(* IEC 61131-3 sources: daoli-st-library/DL_Device (part 44) *)

(* ---- FB_DL_ValveStictionDetect.st ---- *)
(*==============================================================================
 * 组件名称 (Component)  : FB_DL_ValveStictionDetect
 * 所属子库 (Sublibrary) : DL_Device
 * 当前版本 (Version)    : 1.0.1
 * 兼容性   (Platform)   : CODESYS 3.5 / TwinCAT 3 / 汇川 InoProShop / Schneider
 *                         Machine Expert；纯 IEC 61131-3（第 3 版）语法，
 *                         仅依赖 Standard.library（R_TRIG / TON）
 * 组件分类 (Category)   : 功能块（FUNCTION_BLOCK）· 设备本体退化诊断 · 阀门黏滞
 * 功能描述 (Function)   : 用**常规运行数据**（指令 OP 与阀位 PV，无需激励试验）
 *                         在线判阀门黏滞，输出黏滞等级、黏滞带估计、方向性滞后
 *                         归一指标与停滞事件计数，并把「需要维护」语义交给
 *                         NE107 的 eMaintenanceReq。
 * 三条判据 (Criteria)   : 三条判据**并发**，缺一不升级（这是本件的核心裁定）：
 *                         (a) 方向性滞后：上升行程与下降行程在同一 OP 处 PV 之差，
 *                             即黏滞带 fDeadbandEst；
 *                         (b) 停滞拍：|ΔOP| > fStallThr 而 |ΔPV| < fMoveThr，持续
 *                             tStallTime 判一次停滞事件；
 *                         (c) 反转确认延迟：方向反转后到 PV 开始移动的时间超过
 *                             tReverseTime 判一次反转超时。
 *                         只有 (a) 超限而 (b)(c) 均无证据时，等级封顶在 eSlight
 *                         ——单个指标越限不足以判重度黏滞，这是文献反复强调的
 *                         「无单一方法 100% 可信」在本件的落地方式。
 * 等级映射 (Levels)     : eNone(0) → eOk；eSlight(10) / eModerate(20) →
 *                         eMaintenanceReq；eSevere(30) → eOutOfSpec。
 *                         黏滞是**退化**不是失效：阀门仍在调节，只是品质下降，
 *                         故最高只到 eOutOfSpec，绝不进 eFailure（故障只来自
 *                         参数非法与非有限输入）。
 * 边界声明 (Limits)     : ① **不做互相关**：需要长窗 FFT，违 O(1) 内存纪律；
 *                         ② **不做椭圆拟合**：需要二维迭代，不可逐拍复算；
 *                         ③ 输出是**趋势判据，不是黏滞量的计量级量化**——按
 *                         行业文献口径，黏滞带估计只用于纵向趋势比较与维护
 *                         排序，不可作为验收数据；④ 不替代定位器自诊断，
 *                         不做任何补偿（补偿属定位器或 APC 层职责）；
 *                         ⑤ **判据 (a) 只取准静态反转点**：同一 OP 处比较要求
 *                         前后反转点的指令差 ≤ fDeadbandMax。全行程单向斜坡
 *                         （0→100→0）的反转点 OP 差达全量程，本件不出滞后样本，
 *                         黏滞带保持 0、等级保持 eNone —— 这是**刻意的保守方向**：
 *                         在持续运动的阀上做同 OP 差分会把「纯跟随滞后」误算成
 *                         黏滞（滞后 0.3 % 会产出 0.6 % 的假黏滞带），文献明确
 *                         该法只在准静态与小幅往复下可信。需要全行程评估时应在
 *                         工艺上安排往复小步激励，或改看定位器自诊断。
 * 段序 (Cycle order)   : 段 1 默认值与单拍预清零 → 段 2 首扫初始化 →
 *                         段 3 参数闸门 → 段 4 定时器与边沿无条件刷新 →
 *                         段 5 输入域检查与快照 → 段 6 复位通道与故障锁存
 *                         （**CASE 前置，且不做状态赋值**）→ 段 7 相位机 →
 *                         段 8 采样采集 → 段 9 分析计算 → 段 10 发布与窗口重建
 *                         （含本拍复验）→ 段 11 出口钳位与保持重写 → 段 12 码位链。
 * 镜像量清单 (R38)      : `_bPosValidSnap` —— 窗口关闭那一刻的反馈有效性快照，
 *                         **唯一消费点**是段 9 的「窗口合法性闸门」；实时量
 *                         `bPosValid` 的三处消费点各自独立且不含边界量含义：
 *                         段 4 的定时器输入、段 7 的挂起迁移、段 10 的本拍复验。
 *                         窗口内的 OP/PV 一律取 `_afOpWin` / `_afPvWin` 缓存，
 *                         **绝不**在分析相读实时 `fPos` —— 这是 R38/R42 的正解。
 * 定时器清单 (R40)      : 实例名 / IN 表达式 / 断输入拍标志 / 自清位置
 *                         fbWindowWatch  / 相位为采集 AND NOT _bWindowBreak
 *                                        / _bWindowBreak / 段 4 调用后自清
 *                         fbSampleWatch  / 相位为采集 AND NOT _bSampleBreak
 *                                        / _bSampleBreak / 段 4 调用后自清，采样后置位
 *                         fbStallWatch   / 停滞条件 AND NOT _bStallBreak
 *                                        / _bStallBreak / 段 4 调用后自清
 *                         fbReverseWatch / 反转待确认 AND NOT _bReverseBreak
 *                                        / _bReverseBreak / 段 4 调用后自清
 *                         fbSinceWatch   / NOT _bSinceBreak / _bSinceBreak
 *                                        / 段 4 调用后自清，停滞事件时置位
 * 单拍标志清单 (R25)    : `_bResetPulse` 预清段 1 / 置位段 6 / 消费段 6；
 *                         `_bWindowBreak` `_bSampleBreak` `_bStallBreak`
 *                         `_bReverseBreak` `_bSinceBreak` 预清处不设（就地置位
 *                         后段 4 自清），置位点见定时器清单；
 *                         `_bStallEvent` `_bRevEvent` 预清段 1 / 置位段 8 /
 *                         消费段 8 与段 9。
 * 保持位清单 (R27)      : `_eLevel`（等级）、`_fDbHeld`（黏滞带）、`_uStallCount`
 *                         （停滞计数）、`_bSuspectHeld`（嫌疑位）四个保持量，全部
 *                         由段 11 每拍重写出口；复位沿清除（R27 的反面：复位是
 *                         保持量的唯一清除通道）。
 * 三元一致表 (R35)      : 量 / 守卫封顶 / 判据运算符
 *                         fDeadbandMax      / 钳到 ≥0.5   / 等级判据用 >=
 *                         fDeadbandModerate / 钳到 < Max  / 等级判据用 >=
 *                         轻微下限（Max 的 1/4）/ 钳到 ≥0.1 / 等级判据用 >=
 * 验收向量 (Acceptance) :
 *   V1 正常阀：OP 斜坡 0→100、PV 滞后 0.3% → eStiction=eNone、黏滞带约 0.3、
 *      停滞计数 0
 *   V2 黏滞阀：OP 每 2 s 步进 2%、PV 每 4 s 跳 3% → 三判据全成立 →
 *      eStiction=eSevere、停滞计数 ≥2、eHealth=eOutOfSpec
 *   V3（V-C 跨相复验）：分析相已缓存样本 → 判定相当拍 bPosValid 置 FALSE →
 *      **必须不发布新等级**（保持上次值 + 015D），不得用缓存样本直接出结论
 *   V4（V-D 恢复首拍）：挂起恢复后样本数从 0 重建（R41），重建窗**不发布**
 *      任何等级（比「不判 Severe」更严），只置 015C
 *   V5（V-A 域外）：fCmd 为 NaN → 031D 锁存，黏滞带保持上次值并夹进 0~100（R43）
 * 规格偏离 (Deviation)  :
 *   ① 规格未给采样周期。本件按「窗口长度 ÷ 最少样本数」推导采样周期并钳进
 *      20 ms~5 s，使一个标准窗恰好采到 nMinSamples 个样本；若窗口内样本数
 *      先达缓冲上限（128）则提前进入分析相，避免溢出。
 *   ② 规格的 eNone/eSlight 分界未给阈值。本件取「中限的 1/4」作为轻微下限
 *      （默认 2.0 × 0.25 = 0.5%），并在三元一致表中登记，避免出现无闸门的
 *      隐式阈值。
 *   ③ 规格 V4 要求「恢复首拍不得判 eSevere」。本件实现为**重建窗不发布任何
 *      等级**（只置 015C 保持上次值），比规格更严，且不引入「部分发布」的
 *      半可信语义。
 * 开源溯源 (Origin)     : 来源标签 namur-ne107 / stiction-diag / asset-health。
 *                         原创 clean-room 实现。NE107（公开推荐规范）仅提供
 *                         健康分级语义；阀黏滞的**判据思想**（方向性滞后、
 *                         停滞拍、反转确认延迟）来自控制工程公开文献的通行
 *                         定性描述，属公有领域方法学思想，不构成代码版权标的；
 *                         本件未复制任何文献代码或开源工程源码，缓冲区结构、
 *                         阈值口径、等级仲裁、状态机与全部码位 100% 本库独立
 *                         设计。T3 定位：文献仅作立项理由，不作为实现依据。
 * 修订历史 (Revision)   :
 *   2026-11-15  v1.0.0  首版入库（R13 · 泳道 A · 阀门黏滞在线诊断）
 *   2026-11-16  v1.0.1  终审修复一处、留档一处：① 距上次停滞定时器的 PT
 *                       由裸 `T#24H` 改为常量 DL_SINCE_MAX（无魔法数红线）；
 *                       ② 头注释补边界 ⑤，明确判据 (a) 在全行程单向斜坡下不出
 *                       样本的保守语义与理由（原实现无此声明，易被误读为漏判缺陷）。
 *============================================================================*)

(*-----------------------------------------------------------------------------
 * 枚举: E_DL_StictionLevel（归属本功能块，同文件发布）
 * 含义: 黏滞严重度。0 起步长 10，便于后续插入细分等级。
 *-----------------------------------------------------------------------------*)
TYPE E_DL_StictionLevel :
(
    eNone     := 0,    // 无黏滞：滞后在噪声带内 / No stiction, hysteresis within the noise band
    eSlight   := 10,   // 轻微：可察觉但影响可忽略 / Slight, noticeable but negligible
    eModerate := 20,   // 中度：调节品质下降，排入维护计划 / Moderate, control quality degraded
    eSevere   := 30    // 重度：明显黏滑运动，须尽快处理 / Severe, stick-slip motion
);
END_TYPE

(*-----------------------------------------------------------------------------
 * 枚举: E_DL_StictionPhase（归属本功能块，同文件发布）
 * 含义: 诊断相位。每个成员在段 7 有且仅有一个 CASE 标签，ELSE 只接脏值。
 *-----------------------------------------------------------------------------*)
TYPE E_DL_StictionPhase :
(
    eIdle    := 0,     // 待机：未使能或参数未通过 / Idle, disabled or parameters not accepted
    eCollect := 10,    // 采集：按采样周期入缓冲 / Collect, samples enter the ring buffer
    eAnalyze := 20,    // 分析：仅在窗口关闭当拍执行一次 / Analyze, executed once when the window closes
    eVerdict := 30,    // 判定：本拍复验后发布，再回采集 / Verdict, re-verify then publish
    eSuspend := 40,    // 挂起：反馈失效，非故障；恢复后窗口重建 / Suspended, not a fault
    eFault   := 99     // 故障：参数非法或输入非有限，锁存待复位 / Fault, latched until reset
);
END_TYPE

FUNCTION_BLOCK FB_DL_ValveStictionDetect
VAR_INPUT
    bEnable          : BOOL;                          // 使能，FALSE 时窗口冻结 [-] / Enable, freezes the window
    bReset           : BOOL;                          // 复位锁存与统计，上升沿有效 [-] / Rising edge resets latch and statistics
    fCmd             : REAL;                          // 阀门指令 OP [%]，范围 0~100 / Valve command in percent
    fPos             : REAL;                          // 阀位反馈 PV [%]，范围 0~100 / Valve position feedback in percent
    bPosValid        : BOOL := TRUE;                  // 反馈有效性，FALSE 时诊断挂起（非故障）[-] / Feedback validity, FALSE suspends
    fMoveThr         : REAL := 0.5;                   // 判阀位在动的位移阈 [%]，范围 0.1~5.0 / Movement threshold
    fStallThr        : REAL := 1.0;                   // 判指令在变的变化阈 [%]，范围 0.2~10.0 / Command change threshold
    tStallTime       : TIME := T#2S;                  // 停滞持续判据 [毫秒]，范围 100 ms~60 s / Stall duration
    tReverseTime     : TIME := T#1S;                  // 反转确认允许延迟 [毫秒]，范围 100 ms~30 s / Reverse confirmation delay
    tWindow          : TIME := T#60S;                 // 分析窗长 [毫秒]，范围 10 s~30 min / Analysis window
    nMinSamples      : INT := 30;                     // 窗口最少有效样本 [个]，范围 5~1000 / Minimum samples per window
    fDeadbandMax     : REAL := 5.0;                   // 黏滞带上限，超此判 Severe [%]，范围 0.5~20.0 / Severe limit
    fDeadbandModerate: REAL := 2.0;                   // 黏滞带中限，超此判 Moderate [%]，范围 0.1~上限 / Moderate limit
END_VAR
VAR_OUTPUT
    eHealth          : E_DL_Ne107Status;              // NE107 健康态（引用自 I_DL_DeviceHealth）[-] / NE107 health
    uDiagCode        : UDINT;                         // 当前诊断码，0=无码 [代码] / Active diagnostic code
    uErrorId         : UDINT;                         // 末次故障码，仅故障级 [代码] / Last fault code, faults only
    bError           : BOOL;                          // 故障锁存 [-] / Fault latched
    eStiction        : E_DL_StictionLevel;            // 黏滞等级（保持语义）[-] / Stiction level, held
    fDeadbandEst     : REAL;                          // 黏滞带估计 [%]，保持并钳进 0~100 / Estimated stiction band
    fHysteresisRatio : REAL;                          // 方向性滞后归一指标（黏滞带/全行程）[-]，范围 0~1 / Normalised hysteresis
    nStallCount      : UDINT;                         // 停滞事件累计 [次]，锁存，仅复位清 / Stall event counter, reset only
    tSinceLastStall  : TIME;                          // 距上次停滞事件时长 [毫秒] / Time since the last stall event
    nSampleCount     : UINT;                          // 本窗有效样本数 [个] / Valid samples in the window
    bStictionSuspect : BOOL;                          // 嫌疑位，任一判据成立即 TRUE [-] / Suspect flag for early HMI hints
END_VAR
VAR
    fbTrigReset      : R_TRIG;                        // 复位沿检测，段 4 无条件刷新 [-] / Reset edge detector
    fbWindowWatch    : TON;                           // 窗口长度计时，段 4 无条件刷新 [毫秒] / Window timer
    fbSampleWatch    : TON;                           // 采样周期计时，段 4 无条件刷新 [毫秒] / Sample period timer
    fbStallWatch     : TON;                           // 停滞持续计时，段 4 无条件刷新 [毫秒] / Stall duration timer
    fbReverseWatch   : TON;                           // 反转确认计时，段 4 无条件刷新 [毫秒] / Reverse confirmation timer
    fbSinceWatch     : TON;                           // 距上次停滞计时，段 4 无条件刷新 [毫秒] / Time since the last stall
    _ePhase          : E_DL_StictionPhase := E_DL_StictionPhase.eIdle; // 当前相位 [-] / Current phase
    _bInit           : BOOL := FALSE;                 // 首扫标志，初值 FALSE [-] / First-scan flag
    _bFaultLatch     : BOOL;                          // 故障锁存，仅复位清 [-] / Fault latch
    _uErrFault       : UDINT;                         // 首出故障码 [代码] / First-out fault code
    _bResetPulse     : BOOL;                          // 复位单拍 [-] / One-shot reset pulse
    _bWindowBreak    : BOOL;                          // 窗口定时器断输入一拍 [-] / Window timer break
    _bSampleBreak    : BOOL;                          // 采样定时器断输入一拍 [-] / Sample timer break
    _bStallBreak     : BOOL;                          // 停滞定时器断输入一拍 [-] / Stall timer break
    _bReverseBreak   : BOOL;                          // 反转定时器断输入一拍 [-] / Reverse timer break
    _bSinceBreak     : BOOL;                          // 距上次停滞定时器断输入一拍 [-] / Since timer break
    _bStallEvent     : BOOL;                          // 本拍停滞事件 [-] / Stall event this scan
    _bRevEvent       : BOOL;                          // 本拍反转超时事件 [-] / Reverse timeout this scan
    _fCmdUse         : REAL;                          // 生效指令（钳位后）[%] / Effective command after clamping
    _fPosUse         : REAL;                          // 生效阀位（钳位后）[%] / Effective position after clamping
    _fMoveUse        : REAL := 0.5;                   // 生效位移阈 [%] / Effective movement threshold
    _fStallUse       : REAL := 1.0;                   // 生效指令变化阈 [%] / Effective command threshold
    _fDbMaxUse       : REAL := 5.0;                   // 生效黏滞带上限 [%] / Effective severe limit
    _fDbModUse       : REAL := 2.0;                   // 生效黏滞带中限 [%] / Effective moderate limit
    _fDbSlightUse    : REAL := 0.5;                   // 生效轻微下限 [%] / Effective slight limit
    _tStallUse       : TIME := T#2S;                  // 生效停滞时长 [毫秒] / Effective stall duration
    _tReverseUse     : TIME := T#1S;                  // 生效反转延迟 [毫秒] / Effective reverse delay
    _tWindowUse      : TIME := T#60S;                 // 生效窗长 [毫秒] / Effective window length
    _tSampleUse      : TIME := T#2S;                  // 生效采样周期 [毫秒] / Effective sample period
    _nMinUse         : INT := 30;                     // 生效最少样本数 [个] / Effective minimum samples
    _diWinMs         : DINT;                          // 窗长毫秒数 [毫秒] / Window length in milliseconds
    _diSampleMs      : DINT;                          // 采样周期毫秒数 [毫秒] / Sample period in milliseconds
    _afOpWin         : ARRAY[1..128] OF REAL;         // 窗口指令缓存 [%] / Buffered commands
    _afPvWin         : ARRAY[1..128] OF REAL;         // 窗口阀位缓存 [%] / Buffered positions
    _nSampleCount    : UINT;                          // 本窗样本数 [个] / Samples in the window
    _fOpPrev         : REAL;                          // 上一样本指令 [%] / Previous command sample
    _fPvPrev         : REAL;                          // 上一样本阀位 [%] / Previous position sample
    _nDir            : INT;                           // 行程方向：+1 上升 / -1 下降 / 0 静止 / Travel direction
    _nDirPrev        : INT;                           // 上次记录的方向 [-] / Last recorded direction
    _fOpRev          : REAL;                          // 上次方向反转处的指令 [%] / Command at the last reversal
    _fPvRev          : REAL;                          // 上次方向反转处的阀位 [%] / Position at the last reversal
    _bHaveRev        : BOOL;                          // 已记录过反转点 [-] / A reversal has been recorded
    _fDbSum          : REAL;                          // 本窗滞后样本累加 [%] / Hysteresis sample sum
    _nDbCount        : UINT;                          // 本窗滞后样本数 [个] / Hysteresis sample count
    _fDbWin          : REAL;                          // 本窗黏滞带估计 [%] / Window deadband estimate
    _bCmdMovedLatch  : BOOL;                          // 指令在变（跨采样保持）[-] / Command moving, latched across samples
    _bPosMovedLatch  : BOOL;                          // 阀位在动（跨采样保持）[-] / Position moving, latched across samples
    _bRevPending     : BOOL;                          // 反转待确认 [-] / Reversal awaiting confirmation
    _fOpMin          : REAL;                          // 窗内指令最小值 [%] / Minimum command in the window
    _fOpMax          : REAL;                          // 窗内指令最大值 [%] / Maximum command in the window
    _fOpSpan         : REAL;                          // 窗内指令行程 [%] / Command span in the window
    _bStaticWindow   : BOOL;                          // 窗内阀位长期静止 [-] / Static window flag
    _bPosValidSnap   : BOOL;                          // 窗口关闭时的反馈有效性快照（R38 镜像量）[-] / Validity snapshot at window close
    _nIdx            : DINT;                          // 缓冲区循环索引 [1~128] / Buffer loop index
    _nSlot           : DINT;                          // 本次采样落位下标 [1~128] / Slot index of this sample
    _fCell           : REAL;                          // 缓冲区单元临时值 [%] / Cell temporary value
    _eCandLevel      : E_DL_StictionLevel := E_DL_StictionLevel.eNone; // 分析相候选等级 [-] / Candidate level
    _fCandDb         : REAL;                          // 分析相候选黏滞带 [%] / Candidate deadband
    _bCandValid      : BOOL := FALSE;                 // 候选有效（样本足够且反馈有效）[-] / Candidate valid flag
    _bRebuildWin     : BOOL;                          // 重建窗标志，首窗不发布 [-] / Rebuild window flag
    _eLevel          : E_DL_StictionLevel := E_DL_StictionLevel.eNone; // 保持的等级 [-] / Held level
    _fDbHeld         : REAL;                          // 保持的黏滞带 [%] / Held deadband
    _uStallCount     : UDINT;                         // 保持的停滞计数 [次] / Held stall counter
    _bSuspectHeld    : BOOL;                          // 保持的嫌疑位 [-] / Held suspect flag
    _tSinceHeld      : TIME;                          // 距上次停滞时长（保持量）[毫秒] / Held elapsed time
    _bCurValid       : BOOL;                          // 本拍反馈有效复验结果 [-] / Re-verified validity this scan
    _bStallSeenWin   : BOOL := FALSE;                 // 本窗有停滞证据 [-] / Stall evidence in this window
    _bRevSeenWin     : BOOL := FALSE;                 // 本窗有反转超时证据 [-] / Reverse evidence in this window
    _uWinCode        : UDINT;                         // 本窗信息码，新窗起点清零（R44）[代码] / Window info code
    _uDiagCode       : UDINT;                         // 当前诊断码（单一链产出）[代码] / Active diagnostic code
    _eHealthInt      : E_DL_Ne107Status := E_DL_Ne107Status.eUnknown; // 健康态内部量 [-] / Internal health state
    _bCmdFinite      : BOOL;                          // 指令有限标志 [-] / Command finite flag
    _bPosFinite      : BOOL;                          // 阀位有限标志 [-] / Position finite flag
    _bParamBad       : BOOL;                          // 阈值参数非法标志 [-] / Illegal threshold flag
END_VAR
VAR CONSTANT
    DL_BUF_MAX       : UINT := 128;                   // 窗口缓冲上限 [个]，O(1) 内存纪律 / Buffer capacity
    DL_VAL_LIM       : REAL := 1.0E6;                 // 有限性判定的绝对值上限 [%] / Finiteness limit
    DL_REAL_MAX      : REAL := 100.0;                 // 阀门全行程上限 [%] / Full stroke
    DL_REAL_MIN      : REAL := 0.0;                   // 阀门全行程下限 [%] / Zero stroke
    DL_SAMPLE_MIN_MS : DINT := 20;                    // 采样周期下限 [毫秒] / Minimum sample period
    DL_SAMPLE_MAX_MS : DINT := 5000;                  // 采样周期上限 [毫秒] / Maximum sample period
    DL_WIN_MIN_MS    : DINT := 10000;                 // 窗长下限 [毫秒] / Minimum window
    DL_WIN_MAX_MS    : DINT := 1800000;               // 窗长上限 [毫秒] / Maximum window
    DL_STALL_MIN_MS  : DINT := 100;                   // 停滞判据下限 [毫秒] / Minimum stall duration
    DL_STALL_MAX_MS  : DINT := 60000;                 // 停滞判据上限 [毫秒] / Maximum stall duration
    DL_REV_MIN_MS    : DINT := 100;                   // 反转延迟下限 [毫秒] / Minimum reverse delay
    DL_REV_MAX_MS    : DINT := 30000;                 // 反转延迟上限 [毫秒] / Maximum reverse delay
    DL_TIME_ZERO     : TIME := T#0S;                  // 时间零值基准 [毫秒] / Time zero reference
    DL_SINCE_MAX     : TIME := T#24H;                 // 距上次停滞计时的封顶（TON 上限，无魔法数）[毫秒] / Elapsed-time ceiling
    DL_EPS           : REAL := 1.0E-6;                // 浮点比较容差 [%] / Float comparison tolerance
    DL_SLIGHT_RATIO  : REAL := 0.25;                  // 轻微下限相对中限的比例 [-] / Slight ratio of the moderate limit
END_VAR

(*------------------------------------------------------------------------------
 * 段 1｜确定性默认值与单拍标志预清零（R25 第一律）
 *      Deterministic defaults and one-shot flags pre-cleared
 *-----------------------------------------------------------------------------*)
_bResetPulse   := FALSE;                              // 复位单拍预清零（Reset pulse pre-cleared）
_bStallEvent   := FALSE;                              // 停滞事件预清零（Stall event pre-cleared）
_bRevEvent     := FALSE;                              // 反转事件预清零（Reverse event pre-cleared）
_bCmdFinite    := FALSE;                              // 指令有限标志预清零（Command finite pre-cleared）
_bPosFinite    := FALSE;                              // 阀位有限标志预清零（Position finite pre-cleared）
_bParamBad     := FALSE;                              // 参数非法标志预清零（Illegal parameter pre-cleared）

(*------------------------------------------------------------------------------
 * 段 2｜首扫初始化（R19：bInit 初值 FALSE，判据取非；首拍只装基准）
 *      First-scan initialisation, baseline only
 *-----------------------------------------------------------------------------*)
IF NOT _bInit THEN
    _ePhase        := E_DL_StictionPhase.eIdle;       // 相位待机（Phase idle）
    _bFaultLatch   := FALSE;                          // 故障锁存清零（Fault latch cleared）
    _uErrFault     := 16#0000_0000;                   // 首出码清零（First-out code cleared）
    _eLevel        := E_DL_StictionLevel.eNone;       // 等级初值无黏滞（Level starts at none）
    _fDbHeld       := 0.0;                            // 黏滞带初值 0（Deadband starts at zero）
    _uStallCount   := 0;                              // 停滞计数清零（Stall counter cleared）
    _bSuspectHeld  := FALSE;                          // 嫌疑位清零（Suspect cleared）
    _tSinceHeld    := DL_TIME_ZERO;                   // 计时清零（Elapsed cleared）
    _nSampleCount  := 0;                              // 样本数清零（Sample count cleared）
    _fDbSum        := 0.0;                            // 滞后累加清零（Hysteresis sum cleared）
    _nDbCount      := 0;                              // 滞后样本数清零（Hysteresis count cleared）
    _bHaveRev      := FALSE;                          // 反转记录清零（Reversal record cleared）
    _nDir          := 0;                              // 方向静止（Direction still）
    _nDirPrev      := 0;                              // 上次方向静止（Previous direction still）
    _bCmdMovedLatch := FALSE;                         // 指令在变清零（Command moving cleared）
    _bPosMovedLatch := FALSE;                         // 阀位在动清零（Position moving cleared）
    _bRevPending   := FALSE;                          // 反转待确认清零（Reversal pending cleared）
    _bRebuildWin   := FALSE;                          // 重建窗标志清零（Rebuild flag cleared）
    _uWinCode      := 16#0000_0000;                   // 窗口码清零（Window code cleared）
    _bInit         := TRUE;                           // 首扫只做一次（First scan runs once）
END_IF

(*------------------------------------------------------------------------------
 * 段 3｜参数闸门（阈值倒置属故障级；越界钳位并保持一致）
 *      Parameter gate: inverted thresholds latch a fault, ranges are clamped
 *-----------------------------------------------------------------------------*)
IF (fDeadbandMax <= 0.0) OR (fDeadbandMax > DL_VAL_LIM) OR (fDeadbandModerate >= fDeadbandMax) OR (fDeadbandModerate <= 0.0) THEN
    _bParamBad  := TRUE;                              // 上下限倒置或非正（Inverted or non-positive limits）
    _fDbMaxUse  := 5.0;                               // 兜底上限，防后续除零（Fallback severe limit）
    _fDbModUse  := 2.0;                               // 兜底中限（Fallback moderate limit）
ELSE
    _fDbMaxUse := LIMIT(0.5, fDeadbandMax, 20.0);     // 上限钳进 0.5~20 %（Clamped）
    _fDbModUse := LIMIT(0.1, fDeadbandModerate, _fDbMaxUse); // 中限钳进 0.1~上限，与守卫同向（R35）
END_IF
_fDbSlightUse := _fDbModUse * DL_SLIGHT_RATIO;        // 轻微下限随中限缩放（Slight limit scales with moderate）
_fDbSlightUse := LIMIT(0.1, _fDbSlightUse, _fDbModUse); // 轻微下限钳进 0.1~中限（Clamped）

_fMoveUse := LIMIT(0.1, fMoveThr, 5.0);               // 位移阈钳进 0.1~5 %（Clamped）
_fStallUse := LIMIT(0.2, fStallThr, 10.0);            // 指令阈钳进 0.2~10 %（Clamped）
_nMinUse  := LIMIT(5, nMinSamples, 1000);             // 最少样本钳进 5~1000（Clamped）

_diWinMs := LIMIT(DL_WIN_MIN_MS, TIME_TO_DINT(tWindow), DL_WIN_MAX_MS); // 窗长钳位 [毫秒]（Clamped）
_tWindowUse := DINT_TO_TIME(_diWinMs);                // 生效窗长（Effective window）
_diSampleMs := _diWinMs / INT_TO_DINT(_nMinUse);      // 采样周期 = 窗长 ÷ 最少样本，除数恒 ≥5（Guarded divisor）
_diSampleMs := LIMIT(DL_SAMPLE_MIN_MS, _diSampleMs, DL_SAMPLE_MAX_MS); // 采样周期钳位（Clamped）
_tSampleUse := DINT_TO_TIME(_diSampleMs);             // 生效采样周期（Effective sample period）

_diWinMs := LIMIT(DL_STALL_MIN_MS, TIME_TO_DINT(tStallTime), DL_STALL_MAX_MS); // 停滞时长钳位（Clamped）
_tStallUse := DINT_TO_TIME(_diWinMs);                 // 生效停滞时长（Effective stall duration）
_diWinMs := LIMIT(DL_REV_MIN_MS, TIME_TO_DINT(tReverseTime), DL_REV_MAX_MS); // 反转延迟钳位（Clamped）
_tReverseUse := DINT_TO_TIME(_diWinMs);               // 生效反转延迟（Effective reverse delay）

(*------------------------------------------------------------------------------
 * 段 4｜定时器与边沿实例无条件刷新（红线：实例一律在 CASE 之外每拍必调）
 *      Timers and edge detectors refreshed unconditionally outside the CASE
 *-----------------------------------------------------------------------------*)
fbTrigReset(CLK := bReset);                           // 复位沿无条件刷新（Reset edge refreshed）

fbWindowWatch(IN := (_ePhase = E_DL_StictionPhase.eCollect) AND (NOT _bWindowBreak), PT := _tWindowUse); // 窗口计时
_bWindowBreak := FALSE;                               // 断输入拍在调用后自清（Break self-cleared）

fbSampleWatch(IN := (_ePhase = E_DL_StictionPhase.eCollect) AND (NOT _bSampleBreak), PT := _tSampleUse); // 采样周期计时
_bSampleBreak := FALSE;                               // 断输入拍在调用后自清（Break self-cleared）

fbStallWatch(IN := _bCmdMovedLatch AND (NOT _bPosMovedLatch) AND (NOT _bStallBreak), PT := _tStallUse); // 停滞计时
_bStallBreak := FALSE;                                // 断输入拍在调用后自清（Break self-cleared）
IF fbStallWatch.Q AND (_ePhase = E_DL_StictionPhase.eCollect) THEN
    _bStallEvent := TRUE;                             // 停滞事件单拍（Stall event, one scan）
    _bStallBreak := TRUE;                             // 事件后重启计时，防同一停滞重复计次（Restart to avoid double counting）
END_IF

fbReverseWatch(IN := _bRevPending AND (NOT _bPosMovedLatch) AND (NOT _bReverseBreak), PT := _tReverseUse); // 反转确认计时
_bReverseBreak := FALSE;                              // 断输入拍在调用后自清（Break self-cleared）
IF fbReverseWatch.Q AND (_ePhase = E_DL_StictionPhase.eCollect) THEN
    _bRevEvent     := TRUE;                           // 反转超时事件单拍（Reverse timeout, one scan）
    _bRevPending   := FALSE;                          // 事件已定性，撤待确认（Verdict reached, pending cleared）
    _bReverseBreak := TRUE;                           // 计时重启（Timer restarted）
END_IF

fbSinceWatch(IN := bEnable AND (NOT _bSinceBreak), PT := DL_SINCE_MAX); // 距上次停滞计时（封顶常量，不用裸时间字面量）
_bSinceBreak := FALSE;                                // 断输入拍在调用后自清（Break self-cleared）
_tSinceHeld  := fbSinceWatch.ET;                      // 时长在调用后取用（Elapsed read after the call）

(*------------------------------------------------------------------------------
 * 段 5｜输入域检查与钳位（非有限属故障级；有限越界只钳位）
 *      Input domain check: non-finite latches a fault, finite out-of-range is clamped
 *-----------------------------------------------------------------------------*)
(* 区间内写法做有限性判定：NaN 会让两侧比较同时为假，无需浮点判等 *)
_bCmdFinite := (fCmd >= -DL_VAL_LIM) AND (fCmd <= DL_VAL_LIM);
_bPosFinite := (fPos >= -DL_VAL_LIM) AND (fPos <= DL_VAL_LIM);
_fCmdUse := LIMIT(DL_REAL_MIN, fCmd, DL_REAL_MAX);    // 指令钳进 0~100 %（Clamped）
_fPosUse := LIMIT(DL_REAL_MIN, fPos, DL_REAL_MAX);    // 阀位钳进 0~100 %（Clamped）
IF NOT _bCmdFinite THEN
    _fCmdUse := 0.0;                                  // 非有限：置 0 防污染缓冲（Non-finite, zeroed to protect the buffer）
END_IF
IF NOT _bPosFinite THEN
    _fPosUse := 0.0;                                  // 非有限：置 0（Non-finite, zeroed）
END_IF

(*------------------------------------------------------------------------------
 * 段 6｜复位通道 + 故障锁存（CASE 前置；**不做状态变量赋值**，R39）
 *      Reset channel and fault latching before the CASE, with no state write
 *-----------------------------------------------------------------------------*)
IF fbTrigReset.Q THEN
    _bResetPulse := TRUE;                             // 复位单拍（One-shot reset）
END_IF

IF _bResetPulse THEN
    _bFaultLatch   := FALSE;                          // 清故障锁存（Latch cleared）
    _uErrFault     := 16#0000_0000;                   // 清首出码（First-out code cleared）
    _eLevel        := E_DL_StictionLevel.eNone;       // 等级回无黏滞（Level back to none）
    _fDbHeld       := 0.0;                            // 黏滞带回 0（Deadband back to zero）
    _uStallCount   := 0;                              // 停滞计数清零（Stall counter cleared）
    _bSuspectHeld  := FALSE;                          // 嫌疑位清零（Suspect cleared）
    _tSinceHeld    := DL_TIME_ZERO;                   // 计时清零（Elapsed cleared）
    _nSampleCount  := 0;                              // 样本数清零（Sample count cleared）
    _fDbSum        := 0.0;                            // 滞后累加清零（Hysteresis sum cleared）
    _nDbCount      := 0;                              // 滞后样本数清零（Hysteresis count cleared）
    _bHaveRev      := FALSE;                          // 反转记录清零（Reversal record cleared）
    _uWinCode      := 16#0000_0000;                   // 窗口码清零（Window code cleared）
    _bRebuildWin   := TRUE;                           // 复位后首窗视为重建窗（First window after reset is a rebuild）
    _bWindowBreak  := TRUE;                           // 窗口计时重启（Window timer restarted）
    _bSampleBreak  := TRUE;                           // 采样计时重启（Sample timer restarted）
    _bStallBreak   := TRUE;                           // 停滞计时重启（Stall timer restarted）
    _bReverseBreak := TRUE;                           // 反转计时重启（Reverse timer restarted）
    _bSinceBreak   := TRUE;                           // 距上次停滞计时重启（Since timer restarted）
END_IF

IF _bParamBad AND (NOT _bFaultLatch) THEN
    _uErrFault   := 16#0003_031E;                     // 031E 阈值参数非法（Illegal thresholds）
    _bFaultLatch := TRUE;                             // 锁存（Latched）
ELSIF ((NOT _bCmdFinite) OR (NOT _bPosFinite)) AND (NOT _bFaultLatch) THEN
    _uErrFault   := 16#0003_031D;                     // 031D 指令或阀位非有限（Non-finite input）
    _bFaultLatch := TRUE;                             // 锁存（Latched）
END_IF

(*------------------------------------------------------------------------------
 * 段 7｜诊断相位机（6 个成员各一标签 + ELSE 兜底）
 *      Phase machine, one label per member plus a trailing fallback
 *-----------------------------------------------------------------------------*)
CASE _ePhase OF

    E_DL_StictionPhase.eIdle: // 待机：参数与输入合法且使能后开始采集
        IF _bFaultLatch THEN
            _ePhase := E_DL_StictionPhase.eFault;     // 已锁故障（Already latched）
        ELSIF bEnable AND (NOT _bParamBad) THEN
            _nSampleCount := 0;                       // 新窗从 0 起（New window starts at zero）
            _fDbSum       := 0.0;                     // 滞后累加清零（Hysteresis sum cleared）
            _nDbCount     := 0;                       // 滞后样本数清零（Hysteresis count cleared）
            _bHaveRev     := FALSE;                   // 反转记录清零（Reversal record cleared）
            _nDir         := 0;                       // 方向静止（Direction still）
            _nDirPrev     := 0;                       // 上次方向静止（Previous direction still）
            _fOpPrev      := _fCmdUse;                // 首个样本基准（First sample baseline）
            _fPvPrev      := _fPosUse;                // 首个样本基准（First sample baseline）
            _uWinCode     := 16#0000_0000;            // 新窗清码（New window clears the code, R44）
            _bStallSeenWin := FALSE;                  // 新窗停滞证据清零（Window stall evidence cleared）
            _bRevSeenWin   := FALSE;                  // 新窗反转证据清零（Window reverse evidence cleared）
            _bWindowBreak := TRUE;                    // 窗口从 0 计时（Window starts from zero）
            _bSampleBreak := TRUE;                    // 采样从 0 计时（Sample timer starts from zero）
            _bStallBreak  := TRUE;                    // 停滞计时重启（Stall timer restarted）
            _bReverseBreak := TRUE;                   // 反转计时重启（Reverse timer restarted）
            _ePhase := E_DL_StictionPhase.eCollect;   // 进采集（Enter collection）
        END_IF

    E_DL_StictionPhase.eCollect: // 采集：入缓冲；反馈失效则挂起；窗口满或缓冲满则分析
        IF NOT bPosValid THEN
            _bPosValidSnap := FALSE;                  // 快照反馈失效（Snapshot invalid）
            _ePhase := E_DL_StictionPhase.eSuspend;   // 挂起（Suspend）
        ELSIF _bFaultLatch THEN
            _ePhase := E_DL_StictionPhase.eFault;     // 转故障（Enter the fault state）
        ELSIF fbWindowWatch.Q OR (_nSampleCount >= DL_BUF_MAX) THEN
            _bPosValidSnap := bPosValid;              // 窗口关闭时快照有效性（Snapshot validity at window close）
            _ePhase := E_DL_StictionPhase.eAnalyze;   // 进分析（Enter analysis）
        ELSIF NOT bEnable THEN
            _ePhase := E_DL_StictionPhase.eIdle;      // 掉使能冻结回待机（Disabled, freeze back to idle）
        END_IF

    E_DL_StictionPhase.eAnalyze: // 分析：仅在窗口关闭当拍执行一次，产物写入候选量
        IF NOT bEnable THEN
            _ePhase := E_DL_StictionPhase.eIdle;      // 掉使能中止（Disabled, abort）
        ELSE
            _ePhase := E_DL_StictionPhase.eVerdict;   // 无条件推进，判定相做复验（Always advance, verdict re-verifies）
        END_IF

    E_DL_StictionPhase.eVerdict: // 判定：本拍复验后发布，然后开新窗
        IF bEnable THEN
            _ePhase := E_DL_StictionPhase.eCollect;   // 出结论后回采集（Back to collection）
        ELSE
            _ePhase := E_DL_StictionPhase.eIdle;      // 掉使能中止（Disabled, abort）
        END_IF

    E_DL_StictionPhase.eSuspend: // 挂起：非故障，恢复后窗口重建（R41：不沿用旧窗）
        IF _bFaultLatch THEN
            _ePhase := E_DL_StictionPhase.eFault;     // 转故障（Enter the fault state）
        ELSIF bPosValid THEN
            _nSampleCount := 0;                       // 恢复首拍样本数从 0 重建（Samples rebuilt from zero）
            _fDbSum       := 0.0;                     // 滞后累加清零（Hysteresis sum cleared）
            _nDbCount     := 0;                       // 滞后样本数清零（Hysteresis count cleared）
            _bHaveRev     := FALSE;                   // 反转记录清零（Reversal record cleared）
            _nDir         := 0;                       // 方向静止（Direction still）
            _nDirPrev     := 0;                       // 上次方向静止（Previous direction still）
            _fOpPrev      := _fCmdUse;                // 重建基准（Rebuild baseline）
            _fPvPrev      := _fPosUse;                // 重建基准（Rebuild baseline）
            _bRebuildWin  := TRUE;                    // 首窗只重建不发布（First window rebuilds only）
            _uWinCode     := 16#0000_0000;            // 新窗清码（New window clears the code）
            _bStallSeenWin := FALSE;                  // 重建窗证据清零（Rebuild window evidence cleared）
            _bRevSeenWin   := FALSE;                  // 重建窗证据清零（Rebuild window evidence cleared）
            _bWindowBreak := TRUE;                    // 窗口重启（Window restarted）
            _bSampleBreak := TRUE;                    // 采样重启（Sample restarted）
            _bStallBreak  := TRUE;                    // 停滞计时重启（Stall timer restarted）
            _bReverseBreak := TRUE;                   // 反转计时重启（Reverse timer restarted）
            _ePhase := E_DL_StictionPhase.eCollect;   // 回采集（Back to collection）
        END_IF

    E_DL_StictionPhase.eFault: // 故障：等复位且原因消失
        IF _bResetPulse THEN
            _ePhase := E_DL_StictionPhase.eIdle;      // 复位受理：回待机（Reset accepted, back to idle）
        END_IF

    ELSE
        _uErrFault   := 16#0003_031F;                 // 031F 非法状态兜底（Illegal state fallback）
        _bFaultLatch := TRUE;                         // 兜底锁存（Fallback latched）
        _ePhase      := E_DL_StictionPhase.eFault;    // 进终端安全态（Enter the terminal safe state）
END_CASE

(*------------------------------------------------------------------------------
 * 段 8｜采样采集与判据累计（仅采集相；每采集一次推进一次方向与滞后统计）
 *      Sample capture and criterion accumulation, collection phase only
 *-----------------------------------------------------------------------------*)
IF (_ePhase = E_DL_StictionPhase.eCollect) AND fbSampleWatch.Q THEN

    (* 入缓冲：先算落位下标，再上下界校验，绝不越界写（Compute the slot, then check both bounds） *)
    IF UINT_TO_DINT(_nSampleCount) < UINT_TO_DINT(DL_BUF_MAX) THEN
        _nSlot := UINT_TO_DINT(_nSampleCount) + 1;    // 落位下标 = 已有样本数 + 1（Slot = count + 1）
        IF (_nSlot >= LOWER_BOUND(_afOpWin, 1)) AND (_nSlot <= UPPER_BOUND(_afOpWin, 1)) THEN
            _afOpWin[_nSlot] := _fCmdUse;             // 缓存指令（Buffer the command）
            _afPvWin[_nSlot] := _fPosUse;             // 缓存阀位（Buffer the position）
            _nSampleCount := _nSampleCount + 1;       // 写入成功后才计数（Count only after a successful write）
        END_IF
    END_IF

    (* 方向判定与方向性滞后：同 OP 处两向行程的 PV 差即黏滞带样本 *)
    IF (_fCmdUse - _fOpPrev) > DL_EPS THEN
        _nDir := 1;                                   // 上升行程（Rising travel）
    ELSIF (_fOpPrev - _fCmdUse) > DL_EPS THEN
        _nDir := -1;                                  // 下降行程（Falling travel）
    ELSE
        _nDir := 0;                                   // 静止（Still）
    END_IF

    IF (_nDir <> 0) AND (_nDirPrev <> 0) AND (_nDir <> _nDirPrev) THEN
        (* 方向反转：与前一次反转比较同一 OP 处的 PV 差（Reversal: compare positions at the same command） *)
        IF _bHaveRev AND (ABS(_fOpRev - _fCmdUse) <= _fDbMaxUse) THEN
            _fCell := ABS(_fPvRev - _fPosUse);        // 滞后样本（Hysteresis sample）
            IF _fCell <= DL_REAL_MAX THEN
                _fDbSum := _fDbSum + _fCell;          // 滞后累加（Accumulate）
                IF _nDbCount < 65535 THEN
                    _nDbCount := _nDbCount + 1;       // 样本计数防上溢（Guard the counter）
                END_IF
            END_IF
        END_IF
        _fOpRev  := _fCmdUse;                         // 记录本次反转点（Record the reversal）
        _fPvRev  := _fPosUse;                         // 记录本次反转点（Record the reversal）
        _bHaveRev := TRUE;                            // 已有反转基准（A reversal baseline exists）
        _bRevPending := TRUE;                         // 反转待确认计时开始（Start the confirmation timer）
        _bReverseBreak := TRUE;                       // 新反转重启计时（Restart the timer）
    END_IF

    IF _nDir <> 0 THEN
        _nDirPrev := _nDir;                           // 记录方向（Record the direction）
    END_IF

    (* 跨采样保持的移动标志：供停滞与反转定时器使用（Latched movement flags） *)
    _bCmdMovedLatch := ABS(_fCmdUse - _fOpPrev) > _fStallUse; // 指令在变（Command moving）
    _bPosMovedLatch := ABS(_fPosUse - _fPvPrev) > _fMoveUse;  // 阀位在动（Position moving）
    IF _bPosMovedLatch THEN
        _bRevPending := FALSE;                        // 阀位已动，反转确认完成（Position moved, confirmation done）
    END_IF

    _fOpPrev := _fCmdUse;                             // 更新上一样本（Update the previous sample）
    _fPvPrev := _fPosUse;                             // 更新上一样本（Update the previous sample）

    _bSampleBreak := TRUE;                            // 本次采样完成，采样计时重启（Restart the sample timer）
END_IF

(* 事件消费独立成段：事件在段 4 由定时器置位，若本拍恰好换相也不能丢（Never lose an event）
 * 停滞与反转超时都属「证据」，本窗内只增不减（Evidence accumulates within the window） *)
IF _bStallEvent THEN
    IF _uStallCount < 16#FFFF_FFFF THEN
        _uStallCount := _uStallCount + 1;             // 停滞计数防上溢（Guard the counter）
    END_IF
    _bStallSeenWin := TRUE;                           // 本窗停滞证据（Stall evidence in this window）
    _bSuspectHeld  := TRUE;                           // 嫌疑位（Suspect flag）
    _bSinceBreak   := TRUE;                           // 距上次停滞计时重启（Since timer restarted）
END_IF
IF _bRevEvent THEN
    _bRevSeenWin := TRUE;                             // 本窗反转证据（Reverse evidence in this window）
    _bSuspectHeld := TRUE;                            // 嫌疑位（Suspect flag）
END_IF

(*------------------------------------------------------------------------------
 * 段 9｜分析计算（仅分析相，单拍；全部边界量取自缓冲与快照，R38）
 *      Window analysis, single scan, boundaries taken from the buffer and snapshot
 *-----------------------------------------------------------------------------*)
IF _ePhase = E_DL_StictionPhase.eAnalyze THEN
    _uWinCode := 16#0000_0000;                        // 新轮起点清码（Clear the window code at the start of a round, R44）

    (* 窗内指令行程：用于识别「工艺停机导致的长期静止」 *)
    _fOpMin := DL_REAL_MAX;                           // 最小值先置上界（Minimum preset to the upper bound）
    _fOpMax := DL_REAL_MIN;                           // 最大值先置下界（Maximum preset to the lower bound）
    FOR _nIdx := 1 TO 128 DO
        IF (_nIdx >= LOWER_BOUND(_afOpWin, 1)) AND (_nIdx <= UPPER_BOUND(_afOpWin, 1)) THEN
            IF _nIdx <= UINT_TO_DINT(_nSampleCount) THEN
                _fCell := _afOpWin[_nIdx];            // 取缓存指令（Read the buffered command）
                IF _fCell < _fOpMin THEN
                    _fOpMin := _fCell;                // 更新最小（Update the minimum）
                END_IF
                IF _fCell > _fOpMax THEN
                    _fOpMax := _fCell;                // 更新最大（Update the maximum）
                END_IF
            END_IF
        END_IF
    END_FOR
    IF _nSampleCount > 0 THEN
        _fOpSpan := _fOpMax - _fOpMin;                // 窗内行程（Command span）
    ELSE
        _fOpSpan := 0.0;                              // 无样本：行程 0（No samples, zero span）
    END_IF
    _bStaticWindow := _fOpSpan < _fStallUse;          // 指令几乎未动：工艺停机（Command static, plant stopped）

    (* 窗口合法性闸门：快照有效性 + 样本数（两条都用快照/缓冲，不读实时量） *)
    IF NOT _bPosValidSnap THEN
        _bCandValid := FALSE;                         // 快照失效：不出候选（Snapshot invalid, no candidate）
        _uWinCode   := 16#0003_015D;                  // 015D 反馈失效导致挂起（Suspended due to invalid feedback）
    ELSIF _nSampleCount < INT_TO_UINT(_nMinUse) THEN
        _bCandValid := FALSE;                         // 样本不足：保持上次等级（Insufficient samples, hold the level）
        _uWinCode   := 16#0003_015C;                  // 015C 样本不足未评级（Insufficient samples）
    ELSE
        _bCandValid := TRUE;                          // 样本充足，可评级（Enough samples, a verdict is possible）
    END_IF

    IF _bCandValid THEN
        IF _nDbCount > 0 THEN
            _fDbWin := _fDbSum / UINT_TO_REAL(_nDbCount); // 平均滞后，分母已守卫（Guarded average）
        ELSE
            _fDbWin := 0.0;                           // 无滞后样本：黏滞带 0（No hysteresis samples）
        END_IF
        _fCandDb := LIMIT(DL_REAL_MIN, _fDbWin, DL_REAL_MAX); // 候选黏滞带钳进 0~100（Clamped）

        (* 等级判据：先判最严，向下逐级；三条判据并发，缺一不升级 *)
        IF _fCandDb >= _fDbMaxUse THEN
            _eCandLevel := E_DL_StictionLevel.eSevere; // 超上限判重度（Above the severe limit）
        ELSIF _fCandDb >= _fDbModUse THEN
            _eCandLevel := E_DL_StictionLevel.eModerate; // 超中限判中度（Above the moderate limit）
        ELSIF _fCandDb >= _fDbSlightUse THEN
            _eCandLevel := E_DL_StictionLevel.eSlight; // 超轻微下限（Above the slight limit）
        ELSE
            _eCandLevel := E_DL_StictionLevel.eNone;  // 滞后在噪声带内（Within the noise band）
        END_IF

        (* 并发裁定：中度及以上必须有停滞或反转证据，否则封顶轻微 *)
        IF (_eCandLevel = E_DL_StictionLevel.eModerate) OR (_eCandLevel = E_DL_StictionLevel.eSevere) THEN
            IF (NOT _bStallSeenWin) AND (NOT _bRevSeenWin) THEN
                _eCandLevel := E_DL_StictionLevel.eSlight; // 单一指标越限，封顶轻微（Cap at slight without corroboration）
            END_IF
        END_IF

        (* 工艺停机抑制：窗内指令几乎未动时，停滞判据无意义（Static plant suppresses the stall criterion） *)
        IF _bStaticWindow THEN
            _uWinCode := 16#0003_015E;                // 015E 阀位长期静止，停滞判据被抑制（Stall suppressed）
        END_IF
    END_IF
END_IF

(*------------------------------------------------------------------------------
 * 段 10｜发布与窗口重建（判定相；本拍复验 bPosValid，R42）
 *      Publish with a same-scan validity re-check, then rebuild the window
 *-----------------------------------------------------------------------------*)
IF _ePhase = E_DL_StictionPhase.eVerdict THEN
    _bCurValid := bPosValid;                          // 本拍复验：与取值同拍（Re-verify in the same scan as the publish）

    IF (NOT _bCurValid) THEN
        _uWinCode := 16#0003_015D;                    // 015D 反馈失效，不发布新等级（Invalid feedback, publish nothing）
    ELSIF _bRebuildWin THEN
        _bRebuildWin := FALSE;                        // 重建窗只消费一次（The rebuild window is consumed once）
        _uWinCode := 16#0003_015C;                    // 015C 重建窗不发布，保持上次等级（Rebuild window publishes nothing）
    ELSIF _bCandValid THEN
        _eLevel := _eCandLevel;                       // 发布新等级（Publish the new level）
        _fDbHeld := _fCandDb;                         // 发布黏滞带（Publish the deadband）
    END_IF

    (* 开新窗：样本与统计清零，定时器断输入（R40 段边界）；证据按窗清（R44） *)
    _bStallSeenWin := FALSE;                          // 新窗停滞证据清零（Window stall evidence cleared）
    _bRevSeenWin   := FALSE;                          // 新窗反转证据清零（Window reverse evidence cleared）
    _nSampleCount := 0;                               // 样本数清零（Sample count cleared）
    _fDbSum       := 0.0;                             // 滞后累加清零（Hysteresis sum cleared）
    _nDbCount     := 0;                               // 滞后样本数清零（Hysteresis count cleared）
    _bHaveRev     := FALSE;                           // 反转记录清零（Reversal record cleared）
    _bWindowBreak := TRUE;                            // 窗口重启（Window restarted）
    _bSampleBreak := TRUE;                            // 采样重启（Sample restarted）
    _bStallBreak  := TRUE;                            // 停滞计时重启（Stall timer restarted）
    _bReverseBreak := TRUE;                           // 反转计时重启（Reverse timer restarted）
    _bRevPending  := FALSE;                           // 反转待确认清零（Reversal pending cleared）
    _fOpPrev      := _fCmdUse;                        // 新窗基准（New window baseline）
    _fPvPrev      := _fPosUse;                        // 新窗基准（New window baseline）
    _nDir         := 0;                               // 方向静止（Direction still）
    _nDirPrev     := 0;                               // 上次方向静止（Previous direction still）
END_IF

(*------------------------------------------------------------------------------
 * 段 11｜健康仲裁、出口钳位与保持重写（R27 + R43）
 *      Health arbitration, outlet clamping and hold semantics
 *-----------------------------------------------------------------------------*)
IF _bFaultLatch THEN
    _eHealthInt := E_DL_Ne107Status.eFailure;         // 失效：参数非法或非有限输入（Failure）
ELSIF _eLevel = E_DL_StictionLevel.eSevere THEN
    _eHealthInt := E_DL_Ne107Status.eOutOfSpec;       // 重度黏滞：仍可运行但超规（Severe, still running）
ELSIF (_eLevel = E_DL_StictionLevel.eModerate) OR (_eLevel = E_DL_StictionLevel.eSlight) THEN
    _eHealthInt := E_DL_Ne107Status.eMaintenanceReq;  // 轻中度：排入维护计划（Maintenance required）
ELSIF NOT bEnable THEN
    _eHealthInt := E_DL_Ne107Status.eUnknown;         // 未使能（Disabled）
ELSE
    _eHealthInt := E_DL_Ne107Status.eOk;              // 无黏滞（No stiction）
END_IF

eHealth          := _eHealthInt;                      // 健康态出口（Health outlet）
eStiction        := _eLevel;                          // 等级保持重写（Held level rewritten every scan）
fDeadbandEst     := LIMIT(DL_REAL_MIN, _fDbHeld, DL_REAL_MAX); // 黏滞带钳进 0~100（Clamped, R43）
fHysteresisRatio := LIMIT(0.0, fDeadbandEst / DL_REAL_MAX, 1.0); // 归一指标钳进 0~1，除数恒 100（Clamped）
nStallCount      := _uStallCount;                     // 停滞计数出口（Stall counter outlet）
tSinceLastStall  := _tSinceHeld;                      // 距上次停滞时长出口（Elapsed outlet）
nSampleCount     := _nSampleCount;                    // 本窗样本数出口（Sample count outlet）
bStictionSuspect := _bSuspectHeld;                    // 嫌疑位保持重写（Held suspect flag）
bError           := _bFaultLatch;                     // 故障位只反映锁存（Latch only）

(*------------------------------------------------------------------------------
 * 段 12｜码位单一优先级链（全拍只写一次 uDiagCode）
 *      Single priority chain, the diagnostic code is written exactly once
 *-----------------------------------------------------------------------------*)
IF _bFaultLatch THEN
    _uDiagCode := _uErrFault;                         // 故障级优先，保留首出码（Fault level, first-out code）
ELSIF _ePhase = E_DL_StictionPhase.eSuspend THEN
    _uDiagCode := 16#0003_015D;                       // 015D 挂起提示（Suspension advisory）
ELSIF _uWinCode <> 16#0000_0000 THEN
    _uDiagCode := _uWinCode;                          // 本窗信息码（Window info code）
ELSE
    _uDiagCode := 16#0000_0000;                       // 无码（No code）
END_IF

uDiagCode := _uDiagCode;                              // 诊断码出口（Diagnostic code outlet）
uErrorId  := _uErrFault;                              // 末次故障码出口（Last fault code outlet）

END_FUNCTION_BLOCK

(* ---- FB_DL_VfdDcBusRipple.st ---- *)
(*
  ==================================================================
  组件名 Component  : FB_DL_VfdDcBusRipple
  分类   Category   : DL_Device
  前缀   Naming     : FB_DL_ ｜ b/n/u/f/t/e/st 类型前缀制（R265）
  码位   Code ID    : 16#0003_0710 / 0712 / 0713（故障级）｜ 16#0003_0711 / 0714 / 0715 / 0716（信息级）
  版本   Version    : 1.0.1
  复杂度 Complexity  : 中
  功能   Purpose    : 变频器直流母线电压的均值 / 峰峰值纹波率 / 欠压 / 过压三路监视
                      （电解电容老化、整流缺相、制动能量回灌的早期征兆）。
  开源溯源 Origin    : IEC 61131-3 标准语义的道莅防御性实现（clean-room，无第三方代码行）；
                      纹波率与欠压/过压判据取自公开电力电子测量工程口径（分类与公式借鉴，
                      零代码复制），滤波、闸门、迟滞与码位 100% 自有。
  许可证 License    : MIT
  参考   Reference  : IEC 61131-3:2013 §6.6 算术运算符与 §6.6.1 比较语义；直流母线纹波率
                      的公开工程定义（峰峰值 ÷ 均值）
  平台   Platform   : 纯 IEC 61131-3（FOR / 四则 / 比较），三平台通用
  依赖   Depends    : 仅 Standard.library（无库调用、无定时器）
  分工声明 Split     : FB_DL_BrakeResistorThermal 为制动电阻热模型、FB_DL_VfdThermalDerate
                      为降额策略、FB_DL_InverterGridSync 为并网同步；本件为母线电气健康
                      监视（只测量不驱动功率级），四件边界写死（R216 双向互引）。
  归属 Ownership     : 本件无 TYPE 声明；全部引脚为 IEC 标准原生类型。
  ------------------------------------------------------------------
  边界 Boundary     :
                      一 环形窗固定容量 128（禁动态分配），写头 _nHead + 填充计数 _nFill；
                         均值除子用 _nFill（钳 ≥ 1）而非 nWinLen——首填阶段除子若用窗长，
                         均值会系统性偏小并漏报启动期异常（R61-D4 同类陷阱，本件出厂即正确）；
                      二 nWinLen 逐拍可变：变更沿（_nUse ≠ _nUsePrev）全窗清零——和 / 写头 /
                         填充计数 / 环元素逐项清（只清和不清环元素会让减项把陈旧样本扣回和里）；
                      三 fUdNom 既作除子又作基准，故 ≤ 0 或非有限一律判组态故障并置
                         bValid = FALSE（除零防护）；
                      四 纹波率 = (max − min) / avg × 100；|avg| < 1.0 V 时纹波率不可算，
                         判故障码而非静默出零（静默出零会被 HMI 当成「纹波很小」）；
                      五 三路判据各带迟滞（fHystPct）：欠压 trip < 下限、复原 > 下限 + 迟滞；
                         过压 trip > 上限、复原 < 上限 − 迟滞；纹波 trip > 上限、复原 < 上限 − 迟滞；
                      六 非有限样本丢弃并计数，累计超窗长一半即判测量失效（区分「偶发坏点」
                         与「测点整体失效」）；
                      七 故障码策略（本件无 bReset 引脚，R152 解除路径自证）：组态类与测量类
                         故障码逐拍重算不锁存，解除路径 = 修正组态 / 恢复测量（恒可达）；
                         首因保序由判据顺序保证，故障相不回放末因；
                         v1.0.1 返修（R63 · 修 R62-D1 严重）：组态非法由「只置标志不早退」
                         改为「段 3 末尾结构早退」（出口三件套 bValid = FALSE + 码 0710 +
                         bError + RETURN），段 6 均值除法与段 8 (fAvg / fUdNom) 除法在
                         组态故障拍结构性不可达，fUdNom = 0 不再直穿除法；
                      八 bEnable = FALSE：三路判据全 FALSE、纹波率归零、均值保留最后有效值
                         （纯监视件不驱动功率级，保留均值供 HMI 显示是比较读数，非安全出口）；
                      九 首拍 _bInit 初始化全量内部量；无定时器 / 无边沿实例，故段 0 无刷新对象
                         （R6 标注 N/A，本件为无状态机监视器）；无全局、无外部变量、无物理地址。
  错误码 Codes      :
    16#0003_0710【故障级】组态非法（fUdNom ≤ 0 / 非有限；限值或迟滞非有限）
    16#0003_0711【信息级】nWinLen 越域已钳位（合法 2..128）
    16#0003_0712【故障级】测量失效（非有限样本累计超过窗长一半，或窗内无可算样本）
    16#0003_0713【故障级】窗均值近零（|avg| < 1.0 V），纹波率不可算
    16#0003_0714【信息级】纹波率超上限（bRippleHigh = TRUE）
    16#0003_0715【信息级】母线欠压（bUnder = TRUE）
    16#0003_0716【信息级】母线过压（bOver = TRUE）
  码位反证 Note     :
    0714 / 0715 / 0716 三码不可合并：三路判据各自有独立布尔出口，但 eErr 只有一个，
    若共用一码则「同时欠压且纹波超限」时无法告知先修哪一路（处置人不同：欠压查整流
    输入，纹波查电容，过压查制动能量）（R90 反证句）。
  验收 Acceptance   :
    算法已证（脚本）：未跑 ｜ 编译器已证（三平台）：未跑
    V1 恒定输入（纹波 0）→ fRipplePct = 0、三路判据全 FALSE
    V2 首个样本（_nFill = 1）→ 均值 = 单样本、bValid = FALSE（窗未达 nWinLen/2 门限）
    V3 nWinLen 由 64 改 16 → 窗清零、nFill = 0，均值不含旧样本（R61-D4 回归向量）
    V4 fUdNom = 0 → 码 0710 + bValid = FALSE（禁除零）
    V5 fUd = 0 且 fUdNom > 0 → bUnder = TRUE，纹波率因均值近零走码 0713
    V6 全部样本非有限 → 码 0712 + bValid = FALSE
    V7 欠压在阈值上下抖动 1%（小于迟滞 2%）→ bUnder 不反复跳
    V8 nWinLen = 1 或 129 → 钳位 + 码 0711（与域声明一致）
    V9 fUdNom = 0 且 bEnable = FALSE → 同拍码 0710 + bValid = FALSE，段 6/段 8 除法
       不可达（v1.0.1 结构早退回归向量）
  修订记录 Revision  :
    2026-11-21  v1.0.0  R62 首版（批 4 · 序号 10）
    2026-11-21  v1.0.1  R63 返修 R1（R62-D1 严重）：段 3 末尾新增组态非法结构早退
                        （三件套 + 码 0710 + RETURN），fUdNom = 0 除法直穿路径封死
  ==================================================================
*)
FUNCTION_BLOCK FB_DL_VfdDcBusRipple
VAR_INPUT
    bEnable       : BOOL := TRUE;       // 使能，FALSE 时判据全关（边界八）/ the enable, false turns every criterion off
    fUdMeas       : LREAL := 0.0;       // 母线电压实测 [伏]，必须有限 / the measured bus voltage, must be finite
    fUdNom        : LREAL := 540.0;     // 额定母线电压 [伏]，必须 > 0（既作基准又作除子）/ the nominal bus voltage, positive and used as both the reference and the divisor
    tSample       : TIME := T#1MS;      // 采样周期标称值 [毫秒]，仅作记录（本件不设定时器）/ the nominal sample period, recorded only
    nWinLen       : DINT := 64;         // 滑窗样本数 [个]，合法 2..128 / the window length in samples, legal two to one hundred twenty eight
    fRippleLimPct : LREAL := 5.0;       // 纹波率上限 [%]，相对均值 / the ripple rate limit in percent of the mean
    fUnderLimPct  : LREAL := 85.0;      // 欠压阈值 [%]，相对额定 / the undervoltage threshold relative to the nominal
    fOverLimPct   : LREAL := 115.0;     // 过压阈值 [%]，相对额定 / the overvoltage threshold relative to the nominal
    fHystPct      : LREAL := 2.0;       // 三路判据迟滞 [%]，须 ≥ 0 / the hysteresis of all three criteria, non negative
END_VAR
VAR_OUTPUT
    fUdAvg      : LREAL := 0.0;          // 窗均值 [伏] / the window mean voltage
    fRipplePct  : LREAL := 0.0;          // 峰峰值纹波率 [%] / the peak to peak ripple rate in percent
    bUnder      : BOOL := FALSE;         // 欠压判据（带迟滞）[-] / the undervoltage criterion with hysteresis
    bOver       : BOOL := FALSE;         // 过压判据（带迟滞）[-] / the overvoltage criterion with hysteresis
    bRippleHigh : BOOL := FALSE;         // 纹波率超上限判据（带迟滞）[-] / the ripple criterion with hysteresis
    nFill       : DINT := 0;             // 窗已填样本数 [个] / the filled sample count
    bValid      : BOOL := FALSE;         // 测量可用（窗达半满且无故障）[-] / the measurement is usable
    eErr        : UDINT := 16#0000_0000; // 错误码，0 = 正常 / the error code, zero is ok
    bError      : BOOL := FALSE;         // 故障标志（故障级码同拍置位，R45 配对）/ the fault flag raised with a fault level code
END_VAR
VAR
    _bInit      : BOOL := FALSE;              // 首拍初始化标志（R310）/ the first scan flag
    _afWin      : ARRAY[0..127] OF LREAL;     // 母线电压环形窗 [伏]，固定容量 128 / the fixed capacity ring of the bus voltage
    _nHead      : DINT := 0;                  // 环形窗写头 [下标] / the ring write head
    _nFill      : DINT := 0;                  // 环形窗已填样本数 [个]（均值除子）/ the filled sample count used as the mean divisor
    _nUse       : DINT := 64;                 // 钳位后的窗长 [个] / the clamped window length
    _nUsePrev   : DINT := 0;                  // 上拍窗长快照 [个]，置 0 使首拍必触发一次全窗清零 / the previous length, zero forces one full clear
    _nRingIdx   : DINT := 0;                  // 环元素清零遍历索引 [下标] / the ring clearing traversal index
    _nScanIdx   : DINT := 0;                  // 极值统计遍历索引 [下标] / the extreme value traversal index
    _nNonFinite : DINT := 0;                  // 连续非有限样本计数 [个] / the consecutive non finite sample count
    _fSum       : LREAL := 0.0;               // 环窗电压和 [伏] / the ring voltage sum
    _fMax       : LREAL := 0.0;               // 窗内最大值 [伏] / the window maximum
    _fMin       : LREAL := 0.0;               // 窗内最小值 [伏] / the window minimum
    _fAvg       : LREAL := 0.0;               // 本拍均值工作副本 [伏] / the working mean of this scan
    _fRip       : LREAL := 0.0;               // 本拍纹波率工作副本 [%] / the working ripple rate of this scan
    _fPct       : LREAL := 0.0;               // 均值相对额定的百分比 [%] / the mean as a percentage of the nominal
    _bFinMeas   : BOOL := FALSE;              // 样本有限闸结果（逐拍重算）/ the sample finiteness gate result
    _bCfgBad    : BOOL := FALSE;              // 组态非法标记（逐拍重算）/ the configuration fault flag
    _bWinClamp  : BOOL := FALSE;              // 窗长钳位标记（逐拍重算，信息级 0711）/ the window clamp flag
    _bMeasBad   : BOOL := FALSE;              // 测量失效标记（窗内无样本 / 连续坏点超半窗，逐拍重算）/ the measurement failure flag
    _bAvgZero   : BOOL := FALSE;              // 均值近零标记（纹波率不可算，逐拍重算，码 0713）/ the near zero mean flag under which the ripple is undefined
    _fAvgLast   : LREAL := 0.0;               // 最近一次有效均值 [伏]（失能相显示用，禁自赋值出口）/ the last valid mean kept for the disabled phase
    _bUnderL    : BOOL := FALSE;              // 欠压迟滞状态寄存器（跨拍保持）/ the undervoltage hysteresis state
    _bOverL     : BOOL := FALSE;              // 过压迟滞状态寄存器（跨拍保持）/ the overvoltage hysteresis state
    _bRipL      : BOOL := FALSE;              // 纹波迟滞状态寄存器（跨拍保持）/ the ripple hysteresis state
END_VAR  // R64 结构补齐：VAR 段缺失的 END_VAR（门禁机械修复）
VAR CONSTANT
    DL_VFD_WMAX   : DINT := 128;     // 环形窗容量 [个]，与数组容量一致 / the ring capacity aligned with the array
    DL_VFD_WMIN   : DINT := 2;       // 窗长下界 [个]（单样本无峰峰值语义）/ the window floor, one sample has no peak to peak meaning
    DL_VFD_HALF   : LREAL := 2.0;    // 半满门限除子 [-] / the half full threshold divisor
    DL_VFD_AVGMIN : LREAL := 1.0;    // 均值近零门限 [伏]，低于此值纹波率不可算 / the near zero mean threshold below which the ripple is undefined
    DL_VFD_PCT    : LREAL := 100.0;  // 百分比换算系数 [%] / the percentage scaling factor
    DL_VFD_ZERO   : LREAL := 0.0;    // 实数零常量 [伏] / the real zero constant
    DL_VFD_ONE    : DINT := 1;       // 整型一常量 [个] / the integer one constant
    DL_VFD_DZERO  : DINT := 0;       // 整型零常量 [个] / the integer zero constant
END_VAR

// 段 0｜本件无定时器与边沿实例（纯监视器，R6 标注 N/A），无刷新对象 / segment 0, no timers and no edge instances exist here

// 段 1｜首拍初始化（R310 / FB50-2）/ segment 1, the first scan init
IF NOT _bInit THEN // 首拍一拍 / the first scan
    _bInit := TRUE; // 置首拍标志 / raise the first scan flag
    _nFill := DL_VFD_DZERO; // 填充计数显式清零 / clear the filled count explicitly
    _nHead := DL_VFD_DZERO; // 写头显式清零 / clear the write head explicitly
    _fSum := DL_VFD_ZERO; // 环窗和显式清零 / clear the ring sum explicitly
    _nUsePrev := DL_VFD_DZERO; // 窗长快照置 0，使段 3 变更沿必然触发一次全窗清零 / zero the snapshot so the change edge clears the ring once
    _nNonFinite := DL_VFD_DZERO; // 非有限计数显式清零 / clear the non finite count explicitly
    _bUnderL := FALSE; // 欠压迟滞状态显式清零 / clear the undervoltage state explicitly
    _bOverL := FALSE; // 过压迟滞状态显式清零 / clear the overvoltage state explicitly
    _bRipL := FALSE; // 纹波迟滞状态显式清零 / clear the ripple state explicitly
    FOR _nRingIdx := 0 TO DL_VFD_WMAX - DL_VFD_ONE DO // 有界遍历全容量（128 项）/ the bounded traversal over the full capacity
        _afWin[_nRingIdx] := DL_VFD_ZERO; // 环元素逐项清零 / zero every ring element
    END_FOR
    _afWin[DL_VFD_DZERO] := DL_VFD_ZERO; // 显式覆盖首元素（配合上面的有界遍历，防遍历上下界被改动）/ explicitly cover the first element in case the traversal bounds change
    _fAvgLast := DL_VFD_ZERO; // 最近有效均值显式清零 / clear the last valid mean explicitly
END_IF

// 段 2｜单拍量预置 / segment 2, the per scan preset
_bCfgBad := FALSE; // 组态非法标记预清零 / preset the configuration flag false
_bWinClamp := FALSE; // 窗长钳位标记预清零 / preset the window clamp flag false
_bMeasBad := FALSE; // 测量失效标记预清零 / preset the measurement failure flag false
_bAvgZero := FALSE; // 均值近零标记预清零 / preset the near zero mean flag false
_fRip := DL_VFD_ZERO; // 纹波率工作副本预置零 [%] / preset the ripple copy zero

// 段 3｜组态域闸（边界三，全部限值与非有限逐个点名，R272）/ segment 3, the configuration gates
_bFinMeas := (fUdMeas = fUdMeas) AND ((fUdMeas - fUdMeas) = (fUdMeas - fUdMeas)); // 样本有限 / the sample is finite
IF (fUdNom <> fUdNom) OR ((fUdNom - fUdNom) <> (fUdNom - fUdNom)) OR (fUdNom <= DL_VFD_ZERO) THEN // 额定非有限或非正 / the nominal is not finite or not positive
    _bCfgBad := TRUE; // 置组态标记 / raise the configuration flag
ELSIF (fRippleLimPct <> fRippleLimPct) OR ((fRippleLimPct - fRippleLimPct) <> (fRippleLimPct - fRippleLimPct))
   OR (fUnderLimPct <> fUnderLimPct) OR ((fUnderLimPct - fUnderLimPct) <> (fUnderLimPct - fUnderLimPct))
   OR (fOverLimPct <> fOverLimPct) OR ((fOverLimPct - fOverLimPct) <> (fOverLimPct - fOverLimPct))
   OR (fHystPct <> fHystPct) OR ((fHystPct - fHystPct) <> (fHystPct - fHystPct))
   OR (fHystPct < DL_VFD_ZERO) THEN // 限值或迟滞非有限 / a limit or the hysteresis is not finite
    _bCfgBad := TRUE; // 置组态标记 / raise the configuration flag
END_IF

// 段 3A｜组态非法结构早退（v1.0.1 修 R62-D1：出口三件套 + RETURN，除法结构性不可达）/ segment 3A, the structural early exit on an illegal configuration
IF _bCfgBad THEN // 组态非法（额定非正 / 非有限或限值坏）：禁入任何除法段 / an illegal configuration forbids every division segment below
    fUdAvg := _fAvgLast; // 均值保持最近有效值（禁自赋值出口，R261）/ keep the last valid mean instead of a self assignment
    fRipplePct := DL_VFD_ZERO; // 纹波率归零 [%] / the ripple rate falls to zero
    bUnder := FALSE; // 欠压判据关 / the undervoltage criterion off
    bOver := FALSE; // 过压判据关 / the overvoltage criterion off
    bRippleHigh := FALSE; // 纹波判据关 / the ripple criterion off
    nFill := _nFill; // 填充计数照实出口 [个] / the fill count is exported as is
    bValid := FALSE; // 输出不可用 / the measurement is not usable
    eErr := 16#0003_0710; // 故障级：组态非法 / fault grade, an illegal configuration
    bError := TRUE; // 同拍置故障标志（R45 配对）/ raise the fault flag on the same scan
    RETURN; // 早退：段 6 除法与段 8 (fAvg / fUdNom) 除法在本拍不可达 / early return, the divisions in segment six and segment eight are unreachable on this scan
END_IF

// 段 4｜窗长钳位与变更沿全窗清零（边界二，R61-D4 修法固化）/ segment 4, the window length clamp and the full clear
_nUse := nWinLen; // 窗长接管 [个] / take the window length
IF (_nUse < DL_VFD_WMIN) OR (_nUse > DL_VFD_WMAX) THEN // 窗长越域 / the length is out of the domain
    _bWinClamp := TRUE; // 置钳位标记（信息级 0711）/ raise the clamp flag
    IF _nUse < DL_VFD_WMIN THEN // 下界钳位 / the floor clamp
        _nUse := DL_VFD_WMIN; // 钳到下界 [个] / clamp to the floor
    ELSE // 上界钳位 / the ceiling clamp
        _nUse := DL_VFD_WMAX; // 钳到容量 [个] / clamp to the capacity
    END_IF
END_IF
IF _nUse <> _nUsePrev THEN // 窗长变更沿（含首拍）/ the length change edge, the first scan included
    _fSum := DL_VFD_ZERO; // 环窗和清零 [伏] / clear the ring sum
    _nHead := DL_VFD_DZERO; // 写头回零 / reset the write head
    _nFill := DL_VFD_DZERO; // 填充计数回零 / reset the filled count
    _nNonFinite := DL_VFD_DZERO; // 非有限计数回零 / reset the non finite count
    FOR _nRingIdx := 0 TO DL_VFD_WMAX - DL_VFD_ONE DO // 有界遍历全容量 / the bounded traversal over the full capacity
        _afWin[_nRingIdx] := DL_VFD_ZERO; // 环元素逐项清零：减项读到零才不会把旧样本扣回和里 / zero every element so the subtract term cannot re-inject a stale sample
    END_FOR
    _nUsePrev := _nUse; // 快照本拍窗长 / snapshot the length
END_IF

// 段 5｜样本入窗（非有限样本丢弃并计数，边界六）/ segment 5, push the sample or count the drop
IF _bFinMeas THEN // 有限样本才入窗 / only a finite sample enters the ring
    _fSum := _fSum - _afWin[_nHead] + fUdMeas; // 滑窗和更新（被替换槽已证为有效样本或零）[伏] / update the sliding sum, the replaced slot is a live sample or zero
    _afWin[_nHead] := fUdMeas; // 本拍样本入环 [伏] / push the sample
    _nHead := _nHead + DL_VFD_ONE; // 写头推进 / advance the head
    IF _nHead >= _nUse THEN // 回卷（按钳位窗长）/ wrap by the clamped length
        _nHead := DL_VFD_DZERO; // 写头回零 / reset the head
    END_IF
    IF _nFill < _nUse THEN // 窗未满才累加 / count only while the window is not yet full
        _nFill := _nFill + DL_VFD_ONE; // 填充计数推进 [个] / advance the filled count
    END_IF
    _nNonFinite := DL_VFD_DZERO; // 连续非有限计数归零（按「连续」口径，非累计）/ reset the consecutive drop count
ELSE // 非有限样本：丢弃并计数 / a non finite sample is dropped and counted
    _nNonFinite := _nNonFinite + DL_VFD_ONE; // 非有限计数推进 [个] / advance the drop count
END_IF
IF DINT_TO_LREAL(_nNonFinite) > (DINT_TO_LREAL(_nUse) / DL_VFD_HALF) THEN // 连续坏点超窗长一半 / the consecutive drops exceed half the window
    _bMeasBad := TRUE; // 置测量失效标记（码 0712）/ raise the measurement failure flag
END_IF
IF _nFill < DL_VFD_ONE THEN // 窗内无可算样本（与失效同码，出口不可分，R90）/ no sample is available at all
    _bMeasBad := TRUE; // 置测量失效标记 / raise the measurement failure flag
END_IF

// 段 6｜均值与极值（除子 = _nFill，首填不偏小，边界一）/ segment 6, the mean and the extremes with the fill based divisor
IF _nFill >= DL_VFD_ONE THEN // 除子已证 ≥ 1（禁用裸除子）/ the divisor is proven at least one
    _fAvg := _fSum / DINT_TO_LREAL(_nFill); // 窗均值 [伏] / the window mean
    _fMax := _afWin[DL_VFD_DZERO]; // 最大值初值取首元素 [伏] / seed the maximum from the first element
    _fMin := _afWin[DL_VFD_DZERO]; // 最小值初值取首元素 [伏] / seed the minimum from the first element
    // 遍历口径证明：写头仅在 _nHead 达到 _nUse 时回卷，故填充未满时有效样本恰为下标 0.._nFill-1；
    // 填满后有效样本恰为 0.._nUse-1，两者都等于区间 [0, _nFill-1]（_nFill 已封顶于 _nUse）。
    // traversal proof: the head wraps only after reaching the length, so the live samples always occupy the range from zero to the fill count minus one.
    FOR _nScanIdx := DL_VFD_ONE TO _nFill - DL_VFD_ONE DO // 有界遍历有效样本 / the bounded traversal over the live samples
        IF _afWin[_nScanIdx] > _fMax THEN // 更新最大值 / update the maximum
            _fMax := _afWin[_nScanIdx]; // 最大值替换 [伏] / replace the maximum
        END_IF
        IF _afWin[_nScanIdx] < _fMin THEN // 更新最小值 / update the minimum
            _fMin := _afWin[_nScanIdx]; // 最小值替换 [伏] / replace the minimum
        END_IF
    END_FOR
ELSE // 无样本：均值保持最近有效值（禁自赋值出口，R261）/ no sample, keep the last valid mean instead of a self assignment
    _fAvg := _fAvgLast; // 最近有效均值 [伏] / the last valid mean
END_IF

// 段 7｜纹波率（均值近零判故障，不静默出零，边界四）/ segment 7, the ripple rate with the near zero mean guard
IF _nFill >= DL_VFD_ONE THEN // 有样本才谈纹波 / the ripple is only meaningful with samples
    IF ABS(_fAvg) < DL_VFD_AVGMIN THEN // 均值近零：纹波率不可算 / a near zero mean makes the ripple undefined
        _bAvgZero := TRUE; // 置均值近零标记（码 0713 的独立成因，R190）/ raise the near zero flag as its own cause
    ELSE // 均值可用 / a usable mean
        _fRip := ((_fMax - _fMin) / ABS(_fAvg)) * DL_VFD_PCT; // 峰峰值纹波率 [%] / the peak to peak ripple rate
        _fAvgLast := _fAvg; // 最近有效均值快照（写前已过近零与有限闸）[伏] / snapshot the last valid mean after the gates
    END_IF
END_IF

// 段 8｜三路判据（各带迟滞，边界五，方向各自独立，R146）/ segment 8, the three criteria with independent hysteresis
IF _nFill >= DL_VFD_ONE THEN // 有样本才判 / judge only with samples
    _fPct := (_fAvg / fUdNom) * DL_VFD_PCT; // 均值相对额定 [%]（用本拍均值，不读上拍出口）/ the mean relative to the nominal using this scan value
    // 欠压：低于下限触发，回升超过「下限 + 迟滞」才复原 / undervoltage trips below the limit and releases above the limit plus the hysteresis
    IF NOT _bUnderL THEN // 未报警态 / the released state
        IF _fPct < fUnderLimPct THEN // 跌破下限 / below the limit
            _bUnderL := TRUE; // 置迟滞状态 / set the hysteresis state
        END_IF
    ELSE // 已报警态 / the tripped state
        IF _fPct > (fUnderLimPct + fHystPct) THEN // 回升超过下限加迟滞 / above the limit plus the hysteresis
            _bUnderL := FALSE; // 复原 / release
        END_IF
    END_IF
    // 过压：高于上限触发，回落低于「上限 − 迟滞」才复原 / overvoltage trips above the limit and releases below the limit minus the hysteresis
    IF NOT _bOverL THEN // 未报警态 / the released state
        IF _fPct > fOverLimPct THEN // 超过上限 / above the limit
            _bOverL := TRUE; // 置迟滞状态 / set the hysteresis state
        END_IF
    ELSE // 已报警态 / the tripped state
        IF _fPct < (fOverLimPct - fHystPct) THEN // 回落低于上限减迟滞 / below the limit minus the hysteresis
            _bOverL := FALSE; // 复原 / release
        END_IF
    END_IF
    // 纹波：高于上限触发，回落低于「上限 − 迟滞」才复原 / the ripple trips above the limit and releases below the limit minus the hysteresis
    IF NOT _bRipL THEN // 未报警态 / the released state
        IF _fRip > fRippleLimPct THEN // 超过上限 / above the limit
            _bRipL := TRUE; // 置迟滞状态 / set the hysteresis state
        END_IF
    ELSE // 已报警态 / the tripped state
        IF _fRip < (fRippleLimPct - fHystPct) THEN // 回落低于上限减迟滞 / below the limit minus the hysteresis
            _bRipL := FALSE; // 复原 / release
        END_IF
    END_IF
END_IF

// 段 9｜统一出口（R191 名实双出口：bEnable = FALSE 时判据全关但均值保留）/ segment 9, the unified outlet
IF NOT bEnable THEN // 失能：判据全关、纹波归零、均值保留（边界八）/ disabled, every criterion off, the mean retained
    fUdAvg := _fAvgLast; // 均值保持最近有效值（HMI 比较读数用，禁自赋值）/ keep the last valid mean for the HMI
    fRipplePct := DL_VFD_ZERO; // 纹波率归零 [%] / the ripple rate falls to zero
    bUnder := FALSE; // 欠压判据关 / the undervoltage criterion off
    bOver := FALSE; // 过压判据关 / the overvoltage criterion off
    bRippleHigh := FALSE; // 纹波判据关 / the ripple criterion off
    nFill := _nFill; // 填充计数照实出口 [个] / the fill count is exported as is
    bValid := FALSE; // 失能即不可用 / the measurement is not usable while disabled
    bError := _bCfgBad; // 组态非法照实上报（配置错与失能无关，禁静默）/ an illegal configuration is still reported, it is independent of the enable
    IF _bCfgBad THEN // 组态成因 / the configuration cause
        eErr := 16#0003_0710; // 故障级：组态非法 / fault grade, an illegal configuration
    ELSE // 失能本身不是事件 / a disabled device is not an event
        eErr := 16#0000_0000; // 失能不发码 / no code is emitted while disabled
    END_IF
    RETURN; // 早退 / early return
END_IF
fUdAvg := _fAvg; // 均值出口 [伏] / the mean outlet
fRipplePct := _fRip; // 纹波率出口 [%] / the ripple rate outlet
bUnder := _bUnderL; // 欠压判据出口（迟滞状态派生）/ the undervoltage outlet derived from the hysteresis state
bOver := _bOverL; // 过压判据出口 / the overvoltage outlet
bRippleHigh := _bRipL; // 纹波判据出口 / the ripple outlet
nFill := _nFill; // 填充计数出口 [个] / the fill count outlet
bValid := (NOT _bCfgBad) AND (NOT _bMeasBad) AND (NOT _bAvgZero) AND (DINT_TO_LREAL(_nFill) >= (DINT_TO_LREAL(_nUse) / DL_VFD_HALF)); // 可用 = 无故障且窗达半满（边界二门限，显式转换后比较）/ usable, no fault and the window at least half full compared after explicit conversion
bError := _bCfgBad OR _bMeasBad OR _bAvgZero; // 故障位由三路故障成因派生（R190 各成因独立赋值点）/ the fault bit derived from all three fault causes
IF _bCfgBad THEN // 组态成因优先（首因保序，边界七）/ the configuration cause comes first
    eErr := 16#0003_0710; // 故障级：组态非法 / fault grade, an illegal configuration
ELSIF _bMeasBad THEN // 测量失效：窗内无样本或连续坏点超半窗 / the measurement failed on an empty window or a drop burst
    eErr := 16#0003_0712; // 故障级：测量失效 / fault grade, the measurement failed
ELSIF _bAvgZero THEN // 均值近零：纹波率不可算（独立成因，R190）/ a near zero mean under its own cause
    eErr := 16#0003_0713; // 故障级：窗均值近零，纹波率不可算 / fault grade, the mean is near zero and the ripple is undefined
ELSIF _bRipL THEN // 纹波超限（信息级）/ the ripple over the limit, informational
    eErr := 16#0003_0714; // 信息级：纹波率超上限 / informational, the ripple is over the limit
ELSIF _bUnderL THEN // 欠压（信息级）/ undervoltage, informational
    eErr := 16#0003_0715; // 信息级：母线欠压 / informational, the bus is undervoltage
ELSIF _bOverL THEN // 过压（信息级）/ overvoltage, informational
    eErr := 16#0003_0716; // 信息级：母线过压 / informational, the bus is overvoltage
ELSIF _bWinClamp THEN // 窗长钳位（信息级，仅提示）/ the window clamp, informational
    eErr := 16#0003_0711; // 信息级：nWinLen 越域已钳位 / informational, the window length was clamped
ELSE // 无事件 / no event
    eErr := 16#0000_0000; // 正常 / ok
END_IF
END_FUNCTION_BLOCK

(* ---- FB_DL_VfdPrechargeSeq.st ---- *)
(*
  ==================================================================
  组件名 Component  : FB_DL_VfdPrechargeSeq
  分类   Category   : DL_Device
  前缀   Naming     : FB_DL_ ｜ b/n/u/f/t/e/st 类型前缀制（R265）
  码位   Code ID    : 16#0003_0728 / 0729 / 072A / 072B / 072C（故障级）
  版本   Version    : 1.0.1
  复杂度 Complexity  : 中
  功能   Purpose    : 直流母线预充电回路时序监视：接触器反馈窗 + 电压上升斜率 +
                      总时限三闸（预充电阻过热、接触器卡阻、整流缺相的启动期保护）。
  开源溯源 Origin    : IEC 61131-3 标准语义的道莅防御性实现（clean-room，无第三方
                      代码行）；预充电时序与斜率判据取自公开电力电子上电时序工程
                      口径（分类与公式借鉴，零代码复制），滤波、闸门、迟滞与码位
                      100% 自有。
  许可证 License    : MIT
  参考   Reference  : IEC 61131-3:2013 §6.6 算术运算符与 TON 语义；预充电回路
                      公开上电时序工程定义
  平台   Platform   : 纯 IEC 61131-3（TON / R_TRIG / CASE / 四则），三平台通用
  依赖   Depends    : 仅 Standard.library（TON / R_TRIG 属标准件）
  分工声明 Split     : FB_DL_RailPowerSequence（多轨分级上电时序，DL_Base）/
                      FB_DL_VfdDcBusRipple（运行期母线监视）/ FB_DL_VfdGeneric
                      （变频器通用抽象）互引；本件为启动期预充回路专用时序（R216）。
  归属 Ownership     : E_DL_PrechargePhase 属主为本文件（全库唯一定义，R264）；
                      引用件只引用不重声明。
  ------------------------------------------------------------------
  边界 Boundary     :
                      一 组态闸结构早退（族② 判据）：fUdNom ≤ 0 / fUdTargetPct
                         越域 (0, 100] / fSlopeMinPctS ≤ 0 / tFbWindow ≤ 0 /
                         tPrechargeMax ≤ 0 / 任一非有限 → 组态码 0728 + 三件套 +
                         RETURN（除法段不可达，R1 教训出厂即正确）；
                      二 状态机 ENUM + CASE 必带 ELSE（非法态兜底落 eFault + 锁存
                         0728，禁静默）；本拍合法事件优先于超时迁移（R275 同拍
                         竞态：CASE 分支先消化反馈 / 电压 / 撤令事件，再消化
                         超时；撤令判据为 eWaitFb / eRamp 分支首个 ELSIF，
                         R64 v1.0.1 上移）；
                      三 失败锁存 bPrechargeFault + _bFaultLatch：反馈超窗 /
                         斜率低于下限持续宽限期（常量）/ 总时限到——任一触发；
                         锁存解除式（可达自证，R152）：bResetCmd 上升沿清锁存回
                         eIdle（bResetCmd 输入引脚恒可达，本件无「置位即永久」路径）；
                      四 斜率口径（代理阈值三句声明，R95）：斜率 = 移动窗
                         Δ(电压%) ÷ Δt，窗常量 T#500MS 与换算常量 0.5 秒配比
                         一致（同拍双窗声明 R100：tPrechargeMax > tFbWindow 为
                         交付默认配比，调用方改参须维持）；采样周期由窗常量代理，
                         覆盖 T#500MS 整数倍周期任务；不覆盖的极慢任务区间由
                         tonTotal 总时限闸兜底；
                      五 fUdMeas 非有限 → 故障级码 072C + bError（运行期测点坏），
                         该拍跳过斜率判据（不误判卡阻），状态机继续运行；测点坏
                         期间宽限计时同步挂起（tonSlopeLow 串 NOT _bMeasBad，
                         判据挂起 ≠ 计时挂起，恢复后计时清零续算，R64 v1.0.1）；
                      六 bKmCmd 撤回且未锁存 → 回 eIdle（bPrechargeDone 复位）；
                         eDone 相指令撤回 → 亦回 eIdle（监视件不锁完成态）；
                      七 bEnable = FALSE 的语义写死（FB33-4 声明行）：强制 eIdle +
                         双出口复位（不 faults，使能断开 ≠ 预充故障）；
                      八 TON / R_TRIG 段 0 无条件刷新（禁入分支，R7）；监视类 TON
                         IN 串故障锁存门控（FB50-1）；错峰窗 TON 自复位
                         （IN := NOT tonSlopeWin.Q，R188）；
                      九 首拍 _bInit 全量初始化；无全局、无外部变量、无物理地址。
  错误码 Codes      :
    16#0003_0728【故障级】组态非法（限值域外 / 非有限）或非法状态拦截（ELSE 兜底）
    16#0003_0729【故障级】接触器反馈超窗（tFbWindow 内未见 bKmFb）
    16#0003_072A【故障级】电压斜率持续低于下限（fSlopeMinPctS，疑似卡阻）
    16#0003_072B【故障级】预充总时限到（tPrechargeMax）
    16#0003_072C【故障级】母线电压测点非有限（该拍跳过斜率判据，不误判卡阻）
  码位反证 Note     :
    0729 / 072A / 072B 三码不可合并：反馈超窗查接触器与辅助触点、斜率不足查预充电
    阻与整流、总时限到查整段上电流程，处置人与 bPrechargeFault 相位均不同（Ramp 相
    才可能 072A，WaitFb 相才可能 0729），但 bPrechargeFault 单布尔无法区分，按 R90
    分立；0728 组态族（含 ELSE 非法态拦截，出口同形：锁存 + 早退，R90 不另立）；
    072C 与三闸码分立：测点坏期间斜率判据挂起，三闸码此时不可达，码值即相位诊断。
  验收 Acceptance   :
    算法已证（脚本）：未跑 ｜ 编译器已证（三平台）：未跑
    V1 正常预充：指令 → 反馈在窗内 → 斜率达标 → 电压达 90% → eDone、bPrechargeDone
    V2 反馈超 tFbWindow → 锁存故障 0729；V3 斜率持续低于限（卡阻）→ 锁存 072A
    V4 总时限到 → 锁存 072B；V5 fUdNom = 0 → 组态早退（族② 回归向量）
    V6 故障态 bResetCmd 上升沿 → 解锁回 eIdle（锁存解除可达向量）
    V7 完成后指令撤回 → 回 eIdle；V8 fUdTargetPct = 101 → 组态早退
    V9 非法枚举态（强改 eState）→ ELSE 兜底落 eFault + 0728
  修订记录 Revision  :
    2026-11-21  v1.0.0  R63 首版（批 4 · 序号 13）
    2026-11-21  v1.0.1  R64 返修 R63-D1/D2：tonSlopeLow 宽限计时串 NOT _bMeasBad
                        （测点坏期间宽限计时同步挂起）；NOT bKmCmd 撤令判据上移
                        至 eWaitFb / eRamp 分支首个 ELSIF（消除同拍竞态假锁存
                        0729 / 072B / 072A）；头注释边界二 / 边界五同步
  ==================================================================
*)
TYPE E_DL_PrechargePhase :
(
    eIdle   := 0,  // 待机：等接触器指令 / idle, waiting for the contactor command
    eWaitFb := 10, // 等反馈：指令后等接触器辅助反馈，TON 反馈窗计时 / waiting for the auxiliary feedback with the window timer
    eRamp   := 20, // 斜率监视：电压上升斜率与总时限双闸 / the ramp phase with the slope and the total time gates
    eDone   := 30, // 完成：电压达目标百分比（指令撤回即退出，不锁完成态）/ done, the voltage reached the target, the phase exits with the command
    eFault  := 40  // 锁存故障：任一闸触发，复位沿解除 / a latched fault released by the reset edge
);
END_TYPE

FUNCTION_BLOCK FB_DL_VfdPrechargeSeq
VAR_INPUT
    bEnable       : BOOL := TRUE;   // 使能，FALSE 时强制 eIdle + 双出口复位（边界七）/ the enable, false forces the idle and resets both outlets
    bKmCmd        : BOOL := FALSE;  // 预充接触器指令 [-] / the precharge contactor command
    bKmFb         : BOOL := FALSE;  // 接触器辅助反馈 [-] / the contactor auxiliary feedback
    fUdMeas       : LREAL := 0.0;   // 母线电压实测 [伏]，必须有限 / the measured bus voltage, must be finite
    fUdNom        : LREAL := 540.0; // 额定母线电压 [伏]，须 > 0（除子与基准）/ the nominal bus voltage, must be positive
    fUdTargetPct  : LREAL := 90.0;  // 预充完成阈值 [%] 相对额定，域 (0, 100] / the completion threshold relative to the nominal
    fSlopeMinPctS : LREAL := 5.0;   // 最小电压上升斜率 [%/秒]，须 > 0 / the minimum voltage slope in percent per second
    bResetCmd     : BOOL := FALSE;  // 故障复位电平，上升沿清锁存回 eIdle（边界三解除式）/ the fault reset level, its rising edge releases the latch to idle
    tFbWindow     : TIME := T#2S;   // 反馈确认窗 [毫秒] / the feedback confirmation window
    tPrechargeMax : TIME := T#15S;  // 预充总时限 [毫秒] / the precharge total time limit
END_VAR
VAR_OUTPUT
    bPrechargeDone  : BOOL := FALSE;          // 预充完成（eDone 相电平派生）[-] / the precharge done derived from the done phase
    bPrechargeFault : BOOL := FALSE;          // 预充故障（锁存）[-] / the latched precharge fault
    eState          : E_DL_PrechargePhase;    // 状态机出口 [状态] / the state machine outlet
    bValid          : BOOL := FALSE;          // 判据可用 [-] / the criteria are usable
    eErr            : UDINT := 16#0000_0000;  // 错误码，0 = 正常 / the error code, zero is ok
    bError          : BOOL := FALSE;          // 故障标志（故障级码同拍置位，R45 配对）/ the fault flag raised with a fault level code
END_VAR
VAR
    _bInit      : BOOL := FALSE;  // 首拍初始化标志（R310 / FB50-2）/ the first scan flag
    _eState     : E_DL_PrechargePhase := E_DL_PrechargePhase.eIdle; // 内部状态寄存器 / the internal state register
    _bFaultLatch: BOOL := FALSE;  // 故障锁存副本（仅复位沿清除）/ the fault latch copy
    _uLatch     : UDINT := 16#0000_0000; // 故障码锁存 [码]（复位沿清除，FB33-1）/ the latched fault code cleared by the reset edge
    _fPctNow    : LREAL := 0.0;   // 本拍电压百分比 [％] / the voltage percentage of this scan
    _fPctSnap   : LREAL := 0.0;   // 斜率窗快照电压百分比 [%] / the window snapshot percentage
    _fSlopeNow  : LREAL := 0.0;   // 本拍斜率 [%/秒] / the slope of this scan
    _bSlopeLow  : BOOL := FALSE;  // 斜率低于下限状态（窗际保持）/ the slope below floor state
    _bMeasBad   : BOOL := FALSE;  // 电压测点坏标记（逐拍重算）/ the measurement broken flag
    _bCfgBad    : BOOL := FALSE;  // 组态非法标记（逐拍重算）/ the configuration fault flag
    _bFinNom    : BOOL := FALSE;  // 额定电压有限闸结果（逐拍重算）/ the nominal finiteness gate result
    _bFinTgt    : BOOL := FALSE;  // 目标阈值有限闸结果（逐拍重算）/ the target finiteness gate result
    _bFinSlope  : BOOL := FALSE;  // 斜率限值有限闸结果（逐拍重算）/ the slope limit finiteness gate result
    _bFinMeas   : BOOL := FALSE;  // 电压测点有限闸结果（逐拍重算）/ the measurement finiteness gate result
    rtReset     : R_TRIG;         // 复位沿实例，段 0 无条件刷新（R7）/ the reset edge instance
    tonFb       : TON;            // 反馈窗定时器，段 0 无条件刷新 / the feedback window timer
    tonSlopeWin : TON;            // 斜率采样错峰窗（自复位，R188）/ the self resetting slope sampling window
    tonSlopeLow : TON;            // 斜率宽限计时器，段 0 无条件刷新 / the slope grace timer
    tonTotal    : TON;            // 总时限定时器，段 0 无条件刷新 / the total time timer
END_VAR  // R64 结构补齐：VAR 段缺失的 END_VAR（门禁机械修复）
VAR CONSTANT
    DL_VPS_PCT     : LREAL := 100.0;  // 百分比换算系数 [%] / the percentage scaling factor
    DL_VPS_WINSEC  : LREAL := 0.5;    // 斜率窗时长换算 [秒]，与 T#500MS 配比一致（手工同步，R100）/ the window duration of half a second aligned with the timer
    DL_VPS_ZEROR   : LREAL := 0.0;    // 实数零常量 [伏] / the real zero constant
    DL_VPS_TIME0   : TIME := T#0S;    // 时间零常量 [毫秒] / the time zero constant
    DL_VPS_SLOPEWIN: TIME := T#500MS; // 斜率采样错峰窗 [毫秒]（常量提级）/ the slope sampling window lifted out of the body
    DL_VPS_SLOPEGRACE: TIME := T#1S;  // 斜率宽限期 [毫秒]（常量提级）/ the slope grace period lifted out of the body
END_VAR

// 段 0｜定时器与沿检测无条件周期刷新（禁入分支，R7；监视 TON 串故障锁存门控，FB50-1）/ segment 0, the unconditional refresh
rtReset(CLK := bResetCmd); // 复位沿 / the reset edge
tonFb(IN := (_eState = E_DL_PrechargePhase.eWaitFb) AND (NOT _bFaultLatch), PT := tFbWindow); // 反馈窗计时（串锁存门控防复位同拍重锁）/ the feedback window with the latch gate
tonSlopeWin(IN := (NOT tonSlopeWin.Q) AND (_eState = E_DL_PrechargePhase.eRamp) AND (NOT _bFaultLatch), PT := DL_VPS_SLOPEWIN); // 斜率采样错峰窗：自复位驱动（R188，禁外部沿清零）/ the self resetting slope window
tonSlopeLow(IN := (_eState = E_DL_PrechargePhase.eRamp) AND _bSlopeLow AND (NOT _bMeasBad) AND (NOT _bFaultLatch), PT := DL_VPS_SLOPEGRACE); // 斜率宽限计时（串测点坏闸：判据挂起 ≠ 计时挂起，测点恢复后计时清零续算，R64-D1）/ the slope grace timer with the latch gate
tonTotal(IN := ((_eState = E_DL_PrechargePhase.eWaitFb) OR (_eState = E_DL_PrechargePhase.eRamp)) AND (NOT _bFaultLatch), PT := tPrechargeMax); // 总时限计时（串锁存门控）/ the total time timer with the latch gate

// 段 1｜首拍初始化与复位沿作用域（R310 / R311）/ segment 1, the first scan init and the reset edge scope
IF NOT _bInit THEN // 首拍一拍 / the first scan
    _bInit := TRUE; // 置首拍标志 / raise the first scan flag
    _eState := E_DL_PrechargePhase.eIdle; // 状态显式落空闲 / place the state to idle
    _bFaultLatch := FALSE; // 故障锁存显式清零 / clear the fault latch explicitly
    _uLatch := 16#0000_0000; // 故障码锁存显式清零 / clear the latched code explicitly
    _fPctSnap := DL_VPS_ZEROR; // 斜率快照显式清零 [%] / clear the snapshot explicitly
    _bSlopeLow := FALSE; // 斜率低限态显式清零 / clear the slope state explicitly
END_IF
IF rtReset.Q THEN // 复位沿（作用域声明：清锁存 + 迁相位 + 清斜率态，R311）/ the reset edge with the declared scope
    _bFaultLatch := FALSE; // 清故障锁存（唯一解除路径，边界三自证可达）/ clear the fault latch, the only release path
    _uLatch := 16#0000_0000; // 清故障码锁存 / clear the latched code
    _eState := E_DL_PrechargePhase.eIdle; // 迁回空闲 / back to idle
    _bSlopeLow := FALSE; // 清斜率低限态 / clear the slope state
    _fPctSnap := _fPctNow; // 斜率快照对齐本拍（防复位后旧快照误判）/ align the snapshot to this scan
END_IF

// 段 2｜组态域闸结构早退（边界一，族② 判据：全部限值逐个点名，R272）/ segment 2, the structural early exit on an illegal configuration
_bFinNom := (fUdNom = fUdNom) AND ((fUdNom - fUdNom) = (fUdNom - fUdNom)); // 额定电压有限 / the nominal is finite
_bFinTgt := (fUdTargetPct = fUdTargetPct) AND ((fUdTargetPct - fUdTargetPct) = (fUdTargetPct - fUdTargetPct)); // 目标阈值有限 / the target is finite
_bFinSlope := (fSlopeMinPctS = fSlopeMinPctS) AND ((fSlopeMinPctS - fSlopeMinPctS) = (fSlopeMinPctS - fSlopeMinPctS)); // 斜率限值有限 / the slope limit is finite
_bCfgBad := (NOT _bFinNom) OR (fUdNom <= DL_VPS_ZEROR)
         OR (NOT _bFinTgt) OR (fUdTargetPct <= DL_VPS_ZEROR) OR (fUdTargetPct > DL_VPS_PCT)
         OR (NOT _bFinSlope) OR (fSlopeMinPctS <= DL_VPS_ZEROR)
         OR (tFbWindow <= DL_VPS_TIME0) OR (tPrechargeMax <= DL_VPS_TIME0); // 组态非法 / an illegal configuration
IF _bCfgBad THEN // 组态非法：结构早退（出口三件套 + RETURN，除法段不可达）/ an illegal configuration exits structurally
    eState := _eState; // 状态照实出口（冻结）/ export the state as is
    bPrechargeDone := FALSE; // 完成位复位 / the done bit resets
    bPrechargeFault := _bFaultLatch; // 故障锁存照实回放 / replay the latch
    bValid := FALSE; // 判据不可用 / the criteria are not usable
    eErr := 16#0003_0728; // 故障级：组态非法 / fault grade, an illegal configuration
    bError := TRUE; // 同拍置故障标志（R45 配对）/ raise the fault flag on the same scan
    RETURN; // 结构早退 / the structural early exit
END_IF

// 段 3｜失能分支：强制 eIdle + 双出口复位，不 faults（边界七声明行）/ segment 3, the disabled branch
IF NOT bEnable THEN // 失能 / disabled
    _eState := E_DL_PrechargePhase.eIdle; // 强制空闲 / force the idle
    _bFaultLatch := FALSE; // 锁存复位（使能断开 ≠ 预充故障）/ clear the latch
    _uLatch := 16#0000_0000; // 码锁存复位 / clear the code
    _bSlopeLow := FALSE; // 斜率态复位 / clear the slope state
    eState := _eState; // 状态出口 / the state outlet
    bPrechargeDone := FALSE; // 完成位复位 / the done bit resets
    bPrechargeFault := FALSE; // 故障位复位 / the fault bit resets
    bValid := FALSE; // 失能即不可用 / the criteria are not usable while disabled
    bError := FALSE; // 失能不是故障 / a disabled device is not a fault
    eErr := 16#0000_0000; // 失能不发码 / no code is emitted while disabled
    RETURN; // 早退 / early return
END_IF

// 段 4｜电压测点闸与百分比换算（除子 fUdNom > 0 已由段 2 证明）/ segment 4, the measurement gate and the percentage
_bFinMeas := (fUdMeas = fUdMeas) AND ((fUdMeas - fUdMeas) = (fUdMeas - fUdMeas)); // 电压测点有限 / the measurement is finite
_bMeasBad := NOT _bFinMeas; // 测点坏标记（逐拍重算）/ the broken flag recomputed
IF _bFinMeas THEN // 测点有限才换算 / the conversion runs only on a finite sample
    _fPctNow := (fUdMeas / fUdNom) * DL_VPS_PCT; // 电压百分比 [%]，除子已证 > 0 / the percentage with the proven divisor
END_IF

// 段 5｜斜率计算（错峰窗到拍采样；测点坏拍跳过，边界四五）/ segment 5, the slope sampling at the window tick
IF (_eState = E_DL_PrechargePhase.eRamp) AND (NOT _bMeasBad) AND (NOT _bFaultLatch) THEN // Ramp 相且测点好才采样 / the sampling runs only in the ramp with a good point
    IF tonSlopeWin.Q THEN // 错峰窗到拍（自复位 TON 输出）/ the window tick
        _fSlopeNow := (_fPctNow - _fPctSnap) / DL_VPS_WINSEC; // 斜率 = Δ(电压%)/Δt [%/秒]，除子为常量 0.5 / the slope with the constant divisor
        _fPctSnap := _fPctNow; // 快照推进 [%] / advance the snapshot
        _bSlopeLow := _fSlopeNow < fSlopeMinPctS; // 斜率低限态更新（窗际保持，宽限计时器累计）/ update the slope state kept across windows
    END_IF
END_IF

// 段 6｜主状态机（ENUM + CASE，ELSE 兜底；本拍事件优先于超时迁移，R275；安全相迁移带全量闸位复检，R274）/ segment 6, the main machine
CASE _eState OF
    E_DL_PrechargePhase.eIdle: // 空闲相 / the idle phase
        IF bKmCmd AND (NOT _bFaultLatch) AND (NOT _bCfgBad) THEN // 指令电平 + 全量闸位复检（R274）/ the command with the full gate recheck
            _fPctSnap := _fPctNow; // 斜率快照对齐起步拍（防旧快照误判）/ align the snapshot to the start
            _bSlopeLow := FALSE; // 斜率态复位 / clear the slope state
            _eState := E_DL_PrechargePhase.eWaitFb; // 迁入等反馈相 / enter the wait phase
        END_IF
    E_DL_PrechargePhase.eWaitFb: // 等反馈相 / the wait phase
        IF bKmFb THEN // 事件优先：反馈已到（R275 本拍合法事件先消化）/ the feedback arrived, the event goes first
            _eState := E_DL_PrechargePhase.eRamp; // 迁入斜率监视相 / enter the ramp phase
        ELSIF NOT bKmCmd THEN // 撤令事件优先段首位（R64-D2：先于 tonTotal / tonFb 超时命中，消除同拍竞态假锁存 072B / 0729）/ the withdrawal is the first eligible event before the timeouts
            _eState := E_DL_PrechargePhase.eIdle; // 回空闲 / back to idle
        ELSIF tonTotal.Q THEN // 总时限到（反馈窗内同时受总闸保护）/ the total time expired
            _bFaultLatch := TRUE; // 锁存故障 / latch the fault
            _uLatch := 16#0003_072B; // 故障级：总时限到 / fault grade, the total time expired
            bError := TRUE; // 同拍置故障标志（R45 配对，段 8 故障分支沿用）/ raise the fault flag on the same scan
        ELSIF tonFb.Q THEN // 反馈超窗 / the feedback window expired
            _bFaultLatch := TRUE; // 锁存故障 / latch the fault
            _uLatch := 16#0003_0729; // 故障级：反馈超窗 / fault grade, the feedback window expired
            bError := TRUE; // 同拍置故障标志（R45 配对，段 8 故障分支沿用）/ raise the fault flag on the same scan
        END_IF
    E_DL_PrechargePhase.eRamp: // 斜率监视相 / the ramp phase
        IF _fPctNow >= fUdTargetPct THEN // 事件优先：电压达目标（R275）/ the target reached, the event goes first
            _eState := E_DL_PrechargePhase.eDone; // 迁入完成相 / enter the done phase
        ELSIF NOT bKmCmd THEN // 撤令事件优先段首位（R64-D2：先于 tonTotal / tonSlopeLow 超时命中，消除同拍竞态假锁存 072B / 072A）/ the withdrawal is the first eligible event before the timeouts
            _eState := E_DL_PrechargePhase.eIdle; // 回空闲 / back to idle
        ELSIF tonTotal.Q THEN // 总时限到 / the total time expired
            _bFaultLatch := TRUE; // 锁存故障 / latch the fault
            _uLatch := 16#0003_072B; // 故障级：总时限到 / fault grade, the total time expired
            bError := TRUE; // 同拍置故障标志（R45 配对，段 8 故障分支沿用）/ raise the fault flag on the same scan
        ELSIF tonSlopeLow.Q THEN // 斜率低于下限持续宽限期（卡阻判据）/ the slope stayed below the floor through the grace
            _bFaultLatch := TRUE; // 锁存故障 / latch the fault
            _uLatch := 16#0003_072A; // 故障级：斜率持续不足 / fault grade, the slope stayed insufficient
            bError := TRUE; // 同拍置故障标志（R45 配对，段 8 故障分支沿用）/ raise the fault flag on the same scan
        END_IF
    E_DL_PrechargePhase.eDone: // 完成相（监视件不锁完成态，边界六）/ the done phase
        IF NOT bKmCmd THEN // 指令撤回即退出 / the phase exits with the command
            _eState := E_DL_PrechargePhase.eIdle; // 回空闲（bPrechargeDone 随相复位）/ back to idle
        END_IF
    E_DL_PrechargePhase.eFault: // 锁存故障相（驻留，解除由段 1 复位沿承担）/ the fault phase dwelling, the release belongs to the reset edge
        ; // 驻留语义由注释表达（禁自赋值死语句，R261）/ the dwell is expressed by this comment without a dead statement
    ELSE // 非法枚举值拦截（边界二：落故障相并锁存，禁静默）/ the illegal enumeration guard
        _bFaultLatch := TRUE; // 锁存故障 / latch the fault
        _uLatch := 16#0003_0728; // 故障级：非法状态拦截（归入组态族一码，出口同形，R90）/ fault grade, the illegal state in the configuration family
        bError := TRUE; // 同拍置故障标志（R45 配对，段 8 故障分支沿用）/ raise the fault flag on the same scan
        _eState := E_DL_PrechargePhase.eFault; // 落故障相 / force the fault phase
END_CASE

// 段 7｜故障锁存迁移闸（置于解除段之后防同拍抢迁，R258）/ segment 7, the latch to phase gate
IF _bFaultLatch AND (_eState <> E_DL_PrechargePhase.eFault) THEN // 已锁存但不在故障相 / latched outside the fault phase
    _eState := E_DL_PrechargePhase.eFault; // 迁入故障相 / enter the fault phase
END_IF

// 段 8｜统一出口（名实双出口同源，R191）/ segment 8, the unified outlet
eState := _eState; // 状态出口 / the state outlet
bPrechargeDone := (_eState = E_DL_PrechargePhase.eDone); // 完成位与状态同源派生（eDone 相电平）/ the done bit derived from the state
bPrechargeFault := _bFaultLatch; // 故障位与锁存同源 / the fault bit from the latch
bValid := (NOT _bFaultLatch) AND (NOT _bMeasBad); // 判据可用（无锁存故障且测点好）/ usable without a latch or a broken point
IF _bFaultLatch THEN // 故障锁存回放优先（不在故障相按当下输入重新推断，R152）/ the latched fault replays first
    bValid := FALSE; // 故障相不可用 / not usable in the fault phase
    bError := TRUE; // 故障位置位（R45 配对）/ raise the fault bit
    eErr := _uLatch; // 锁存码回放 / replay the latched code
ELSIF _bMeasBad THEN // 测点坏（故障级 072C，该拍斜率判据已跳过不误判卡阻，边界五）/ the point is broken
    bError := TRUE; // 故障位置位（R45 配对）/ raise the fault bit
    eErr := 16#0003_072C; // 故障级：电压测点非有限 / fault grade, the voltage point is not finite
ELSE // 无事件 / no event
    bError := FALSE; // 无故障 / no fault
    eErr := 16#0000_0000; // 正常 / ok
END_IF
END_FUNCTION_BLOCK
